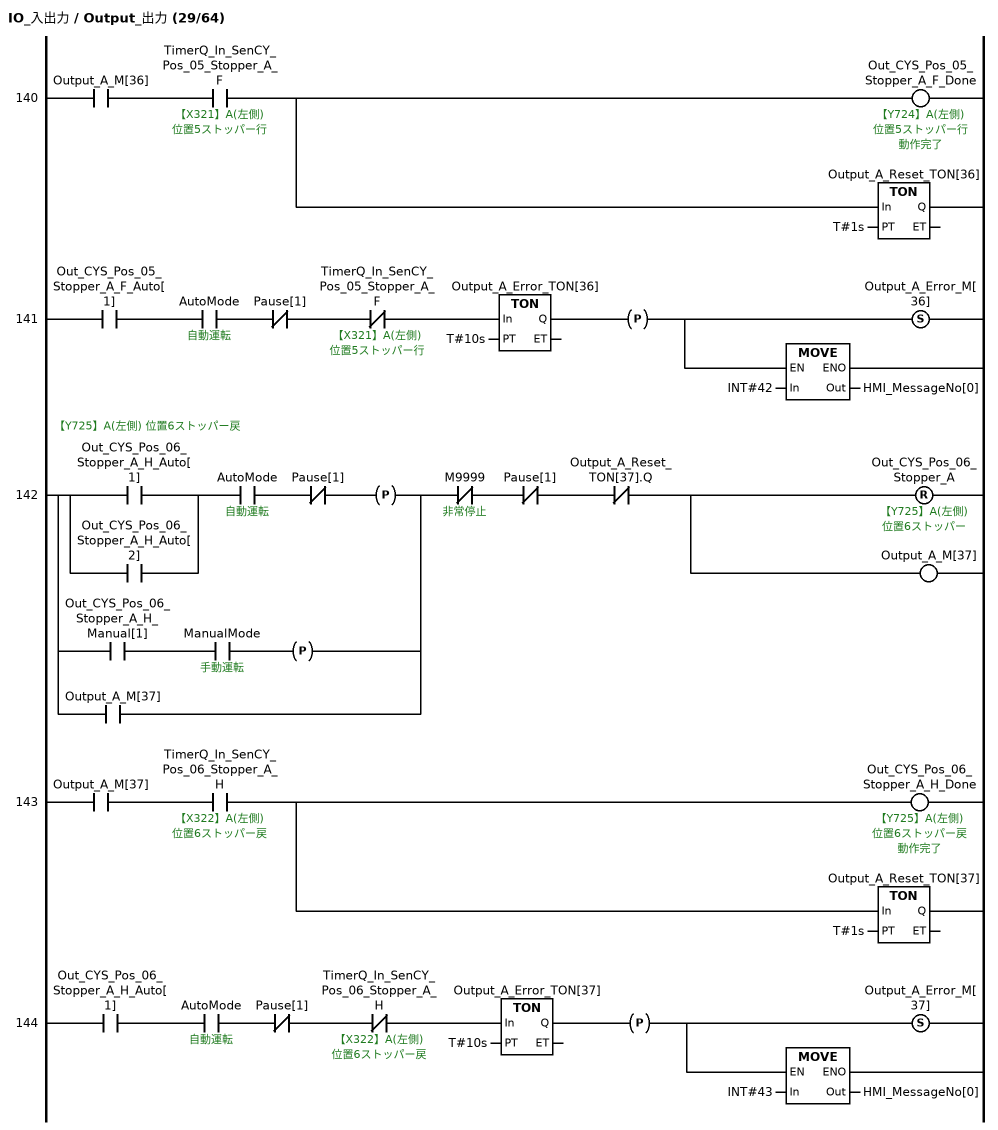
(* [picture p141: IO_入出力 / Output_出力, rungs 140-144] *)
(* Rung 140 *)
_p196 := Output_A_M[36] AND TimerQ_In_SenCY_Pos_05_Stopper_A_F;
Out_CYS_Pos_05_Stopper_A_F_Done := _p196;
Output_A_Reset_TON[36](In := _p196, PT := T#1s);
(* Rung 141 *)
Output_A_Error_TON[36](In := Out_CYS_Pos_05_Stopper_A_F_Auto[1] AND AutoMode AND NOT Pause[1] AND NOT TimerQ_In_SenCY_Pos_05_Stopper_A_F, PT := T#10s);
_e197(CLK := Output_A_Error_TON[36].Q);
IF _e197.Q THEN
    Output_A_Error_M[36] := TRUE;
    HMI_MessageNo[0] := INT#42;
END_IF;
(* Rung 142: 【Y725】A(左側) 位置6ストッパー戻 *)
_e198(CLK := (Out_CYS_Pos_06_Stopper_A_H_Auto[1] OR Out_CYS_Pos_06_Stopper_A_H_Auto[2]) AND AutoMode AND NOT Pause[1]);
_e199(CLK := Out_CYS_Pos_06_Stopper_A_H_Manual[1] AND ManualMode);
_p200 := (_e198.Q OR _e199.Q OR Output_A_M[37]) AND NOT M9999 AND NOT Pause[1] AND NOT Output_A_Reset_TON[37].Q;
IF _p200 THEN Out_CYS_Pos_06_Stopper_A := FALSE; END_IF;
Output_A_M[37] := _p200;
(* Rung 143 *)
_p201 := Output_A_M[37] AND TimerQ_In_SenCY_Pos_06_Stopper_A_H;
Out_CYS_Pos_06_Stopper_A_H_Done := _p201;
Output_A_Reset_TON[37](In := _p201, PT := T#1s);
(* Rung 144 *)
Output_A_Error_TON[37](In := Out_CYS_Pos_06_Stopper_A_H_Auto[1] AND AutoMode AND NOT Pause[1] AND NOT TimerQ_In_SenCY_Pos_06_Stopper_A_H, PT := T#10s);
_e202(CLK := Output_A_Error_TON[37].Q);
IF _e202.Q THEN
    Output_A_Error_M[37] := TRUE;
    HMI_MessageNo[0] := INT#43;
END_IF;

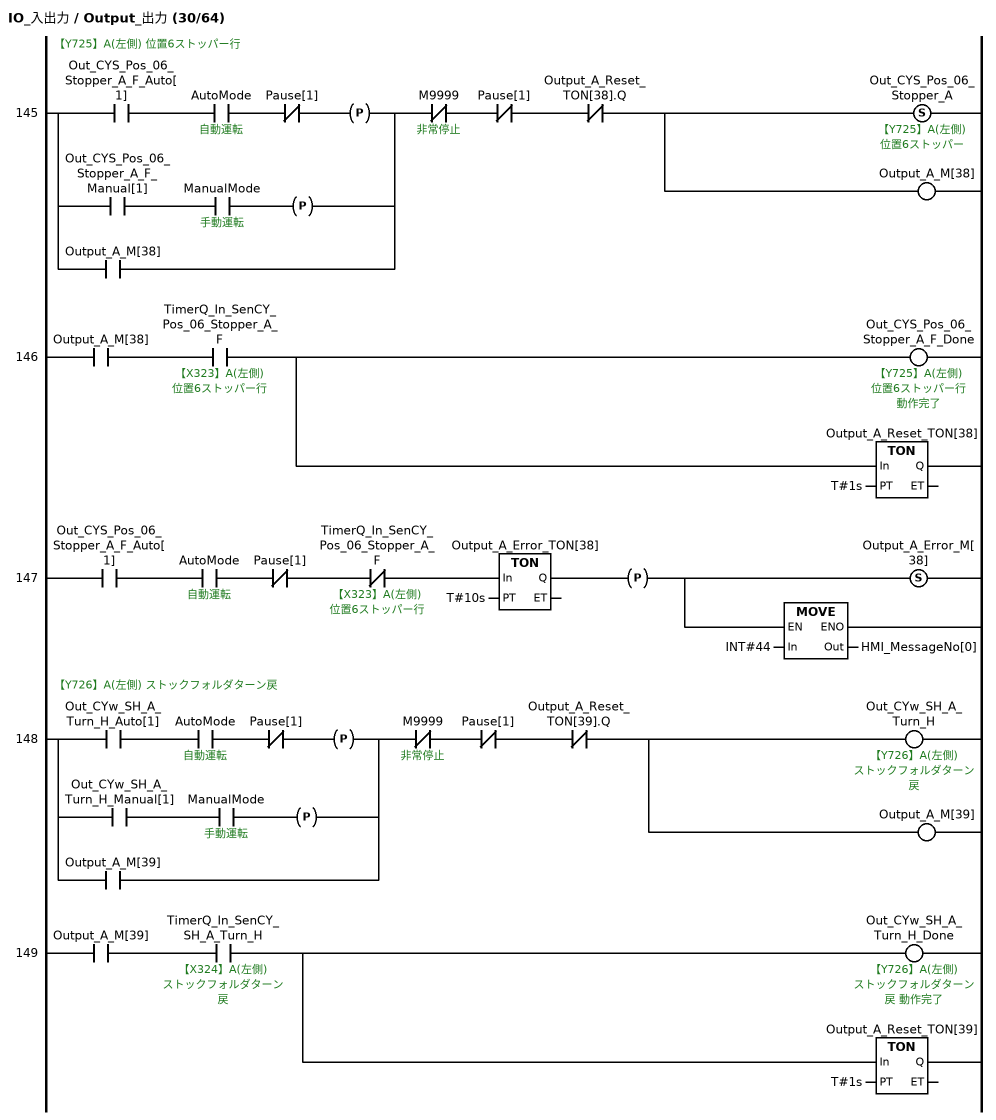
(* Rung 145: 【Y725】A(左側) 位置6ストッパー行 *)
_e203(CLK := Out_CYS_Pos_06_Stopper_A_F_Auto[1] AND AutoMode AND NOT Pause[1]);
_e204(CLK := Out_CYS_Pos_06_Stopper_A_F_Manual[1] AND ManualMode);
_p205 := (_e203.Q OR _e204.Q OR Output_A_M[38]) AND NOT M9999 AND NOT Pause[1] AND NOT Output_A_Reset_TON[38].Q;
IF _p205 THEN Out_CYS_Pos_06_Stopper_A := TRUE; END_IF;
Output_A_M[38] := _p205;
(* Rung 146 *)
_p206 := Output_A_M[38] AND TimerQ_In_SenCY_Pos_06_Stopper_A_F;
Out_CYS_Pos_06_Stopper_A_F_Done := _p206;
Output_A_Reset_TON[38](In := _p206, PT := T#1s);
(* Rung 147 *)
Output_A_Error_TON[38](In := Out_CYS_Pos_06_Stopper_A_F_Auto[1] AND AutoMode AND NOT Pause[1] AND NOT TimerQ_In_SenCY_Pos_06_Stopper_A_F, PT := T#10s);
_e207(CLK := Output_A_Error_TON[38].Q);
IF _e207.Q THEN
    Output_A_Error_M[38] := TRUE;
    HMI_MessageNo[0] := INT#44;
END_IF;
(* Rung 148: 【Y726】A(左側) ストックフォルダターン戻 *)
_e208(CLK := Out_CYw_SH_A_Turn_H_Auto[1] AND AutoMode AND NOT Pause[1]);
_e209(CLK := Out_CYw_SH_A_Turn_H_Manual[1] AND ManualMode);
_p210 := (_e208.Q OR _e209.Q OR Output_A_M[39]) AND NOT M9999 AND NOT Pause[1] AND NOT Output_A_Reset_TON[39].Q;
Out_CYw_SH_A_Turn_H := _p210;
Output_A_M[39] := _p210;
(* Rung 149 *)
Out_CYw_SH_A_Turn_H_Done := Output_A_M[39] AND TimerQ_In_SenCY_SH_A_Turn_H;
Output_A_Reset_TON[39](In := Output_A_M[39] AND TimerQ_In_SenCY_SH_A_Turn_H, PT := T#1s);

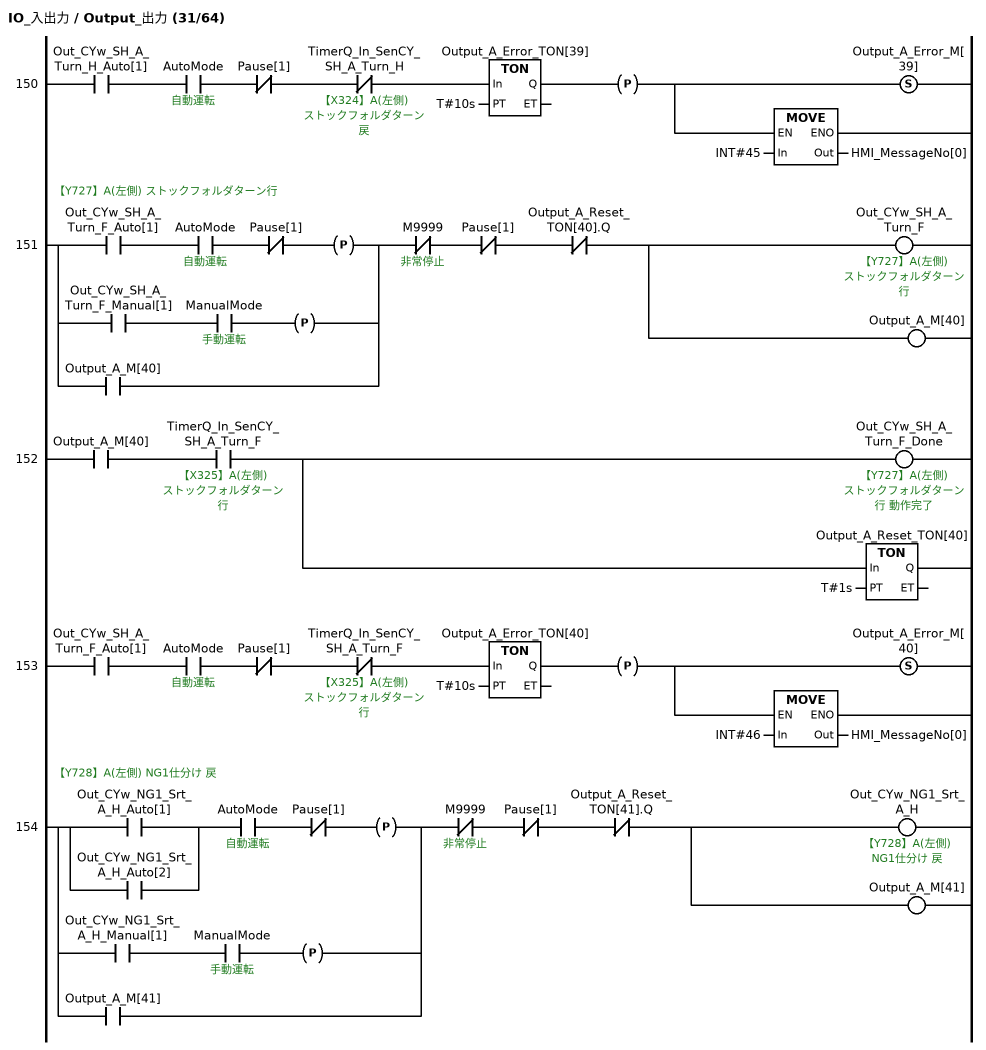
(* Rung 150 *)
Output_A_Error_TON[39](In := Out_CYw_SH_A_Turn_H_Auto[1] AND AutoMode AND NOT Pause[1] AND NOT TimerQ_In_SenCY_SH_A_Turn_H, PT := T#10s);
_e211(CLK := Output_A_Error_TON[39].Q);
IF _e211.Q THEN
    Output_A_Error_M[39] := TRUE;
    HMI_MessageNo[0] := INT#45;
END_IF;
(* Rung 151: 【Y727】A(左側) ストックフォルダターン行 *)
_e212(CLK := Out_CYw_SH_A_Turn_F_Auto[1] AND AutoMode AND NOT Pause[1]);
_e213(CLK := Out_CYw_SH_A_Turn_F_Manual[1] AND ManualMode);
_p214 := (_e212.Q OR _e213.Q OR Output_A_M[40]) AND NOT M9999 AND NOT Pause[1] AND NOT Output_A_Reset_TON[40].Q;
Out_CYw_SH_A_Turn_F := _p214;
Output_A_M[40] := _p214;
(* Rung 152 *)
Out_CYw_SH_A_Turn_F_Done := Output_A_M[40] AND TimerQ_In_SenCY_SH_A_Turn_F;
Output_A_Reset_TON[40](In := Output_A_M[40] AND TimerQ_In_SenCY_SH_A_Turn_F, PT := T#1s);
(* Rung 153 *)
Output_A_Error_TON[40](In := Out_CYw_SH_A_Turn_F_Auto[1] AND AutoMode AND NOT Pause[1] AND NOT TimerQ_In_SenCY_SH_A_Turn_F, PT := T#10s);
_e215(CLK := Output_A_Error_TON[40].Q);
IF _e215.Q THEN
    Output_A_Error_M[40] := TRUE;
    HMI_MessageNo[0] := INT#46;
END_IF;
(* Rung 154: 【Y728】A(左側) NG1仕分け 戻 *)
_e216(CLK := (Out_CYw_NG1_Srt_A_H_Auto[1] OR Out_CYw_NG1_Srt_A_H_Auto[2]) AND AutoMode AND NOT Pause[1]);
_e217(CLK := Out_CYw_NG1_Srt_A_H_Manual[1] AND ManualMode);
_p218 := (_e216.Q OR _e217.Q OR Output_A_M[41]) AND NOT M9999 AND NOT Pause[1] AND NOT Output_A_Reset_TON[41].Q;
Out_CYw_NG1_Srt_A_H := _p218;
Output_A_M[41] := _p218;

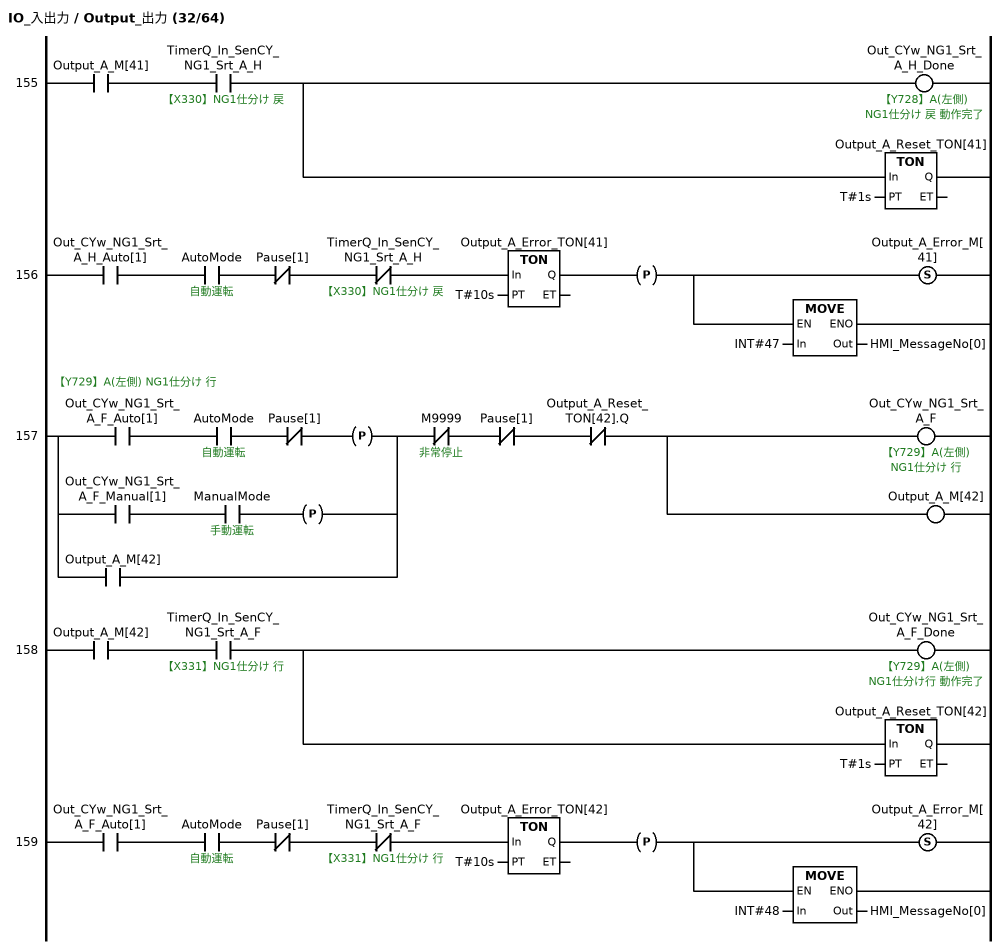
(* Rung 155 *)
Out_CYw_NG1_Srt_A_H_Done := Output_A_M[41] AND TimerQ_In_SenCY_NG1_Srt_A_H;
Output_A_Reset_TON[41](In := Output_A_M[41] AND TimerQ_In_SenCY_NG1_Srt_A_H, PT := T#1s);
(* Rung 156 *)
Output_A_Error_TON[41](In := Out_CYw_NG1_Srt_A_H_Auto[1] AND AutoMode AND NOT Pause[1] AND NOT TimerQ_In_SenCY_NG1_Srt_A_H, PT := T#10s);
_e219(CLK := Output_A_Error_TON[41].Q);
IF _e219.Q THEN
    Output_A_Error_M[41] := TRUE;
    HMI_MessageNo[0] := INT#47;
END_IF;
(* Rung 157: 【Y729】A(左側) NG1仕分け 行 *)
_e220(CLK := Out_CYw_NG1_Srt_A_F_Auto[1] AND AutoMode AND NOT Pause[1]);
_e221(CLK := Out_CYw_NG1_Srt_A_F_Manual[1] AND ManualMode);
_p222 := (_e220.Q OR _e221.Q OR Output_A_M[42]) AND NOT M9999 AND NOT Pause[1] AND NOT Output_A_Reset_TON[42].Q;
Out_CYw_NG1_Srt_A_F := _p222;
Output_A_M[42] := _p222;
(* Rung 158 *)
Out_CYw_NG1_Srt_A_F_Done := Output_A_M[42] AND TimerQ_In_SenCY_NG1_Srt_A_F;
Output_A_Reset_TON[42](In := Output_A_M[42] AND TimerQ_In_SenCY_NG1_Srt_A_F, PT := T#1s);
(* Rung 159 *)
Output_A_Error_TON[42](In := Out_CYw_NG1_Srt_A_F_Auto[1] AND AutoMode AND NOT Pause[1] AND NOT TimerQ_In_SenCY_NG1_Srt_A_F, PT := T#10s);
_e223(CLK := Output_A_Error_TON[42].Q);
IF _e223.Q THEN
    Output_A_Error_M[42] := TRUE;
    HMI_MessageNo[0] := INT#48;
END_IF;

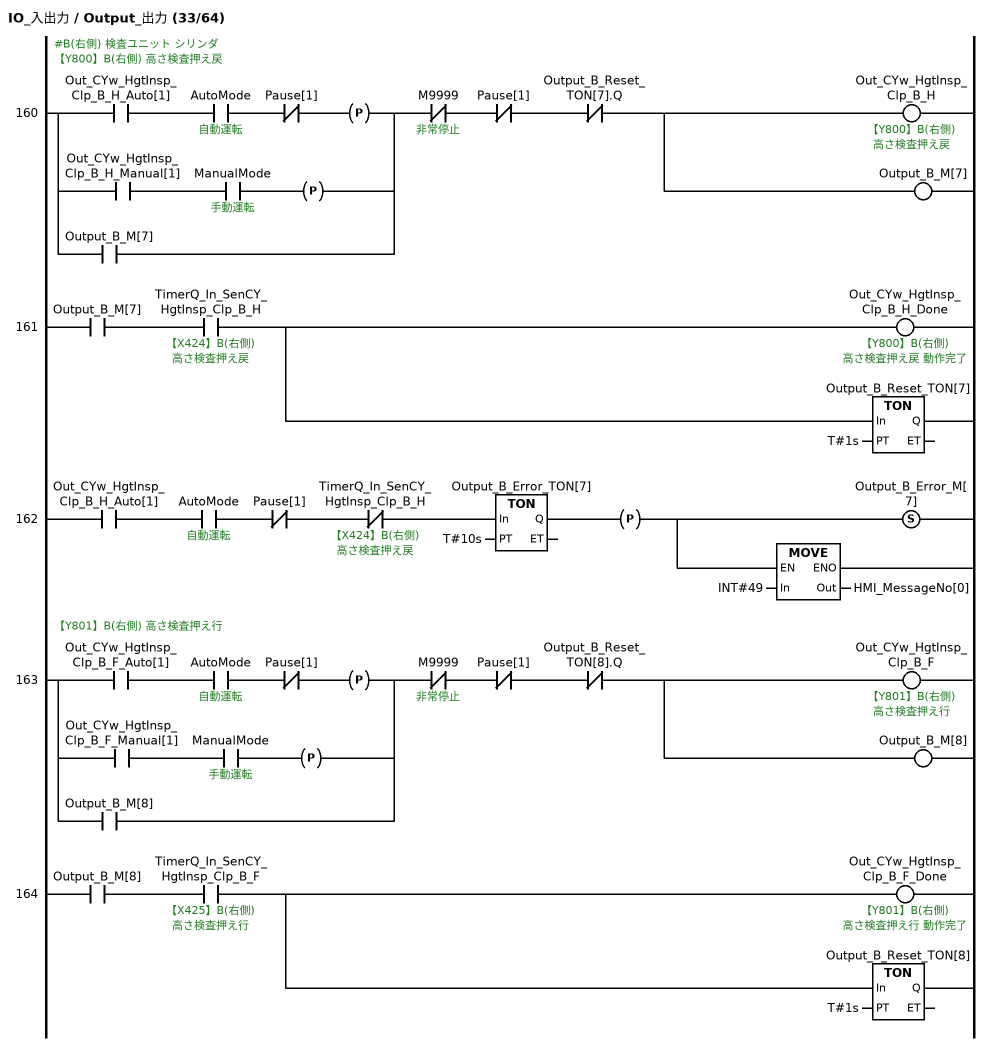
(* Rung 160: #B(右側) 検査ユニット シリンダ / 【Y800】B(右側) 高さ検査押え戻 *)
_e224(CLK := Out_CYw_HgtInsp_Clp_B_H_Auto[1] AND AutoMode AND NOT Pause[1]);
_e225(CLK := Out_CYw_HgtInsp_Clp_B_H_Manual[1] AND ManualMode);
_p226 := (_e224.Q OR _e225.Q OR Output_B_M[7]) AND NOT M9999 AND NOT Pause[1] AND NOT Output_B_Reset_TON[7].Q;
Out_CYw_HgtInsp_Clp_B_H := _p226;
Output_B_M[7] := _p226;
(* Rung 161 *)
_p227 := Output_B_M[7] AND TimerQ_In_SenCY_HgtInsp_Clp_B_H;
Out_CYw_HgtInsp_Clp_B_H_Done := _p227;
Output_B_Reset_TON[7](In := _p227, PT := T#1s);
(* Rung 162 *)
Output_B_Error_TON[7](In := Out_CYw_HgtInsp_Clp_B_H_Auto[1] AND AutoMode AND NOT Pause[1] AND NOT TimerQ_In_SenCY_HgtInsp_Clp_B_H, PT := T#10s);
_e228(CLK := Output_B_Error_TON[7].Q);
IF _e228.Q THEN
    Output_B_Error_M[7] := TRUE;
    HMI_MessageNo[0] := INT#49;
END_IF;
(* Rung 163: 【Y801】B(右側) 高さ検査押え行 *)
_e229(CLK := Out_CYw_HgtInsp_Clp_B_F_Auto[1] AND AutoMode AND NOT Pause[1]);
_e230(CLK := Out_CYw_HgtInsp_Clp_B_F_Manual[1] AND ManualMode);
_p231 := (_e229.Q OR _e230.Q OR Output_B_M[8]) AND NOT M9999 AND NOT Pause[1] AND NOT Output_B_Reset_TON[8].Q;
Out_CYw_HgtInsp_Clp_B_F := _p231;
Output_B_M[8] := _p231;
(* Rung 164 *)
_p232 := Output_B_M[8] AND TimerQ_In_SenCY_HgtInsp_Clp_B_F;
Out_CYw_HgtInsp_Clp_B_F_Done := _p232;
Output_B_Reset_TON[8](In := _p232, PT := T#1s);

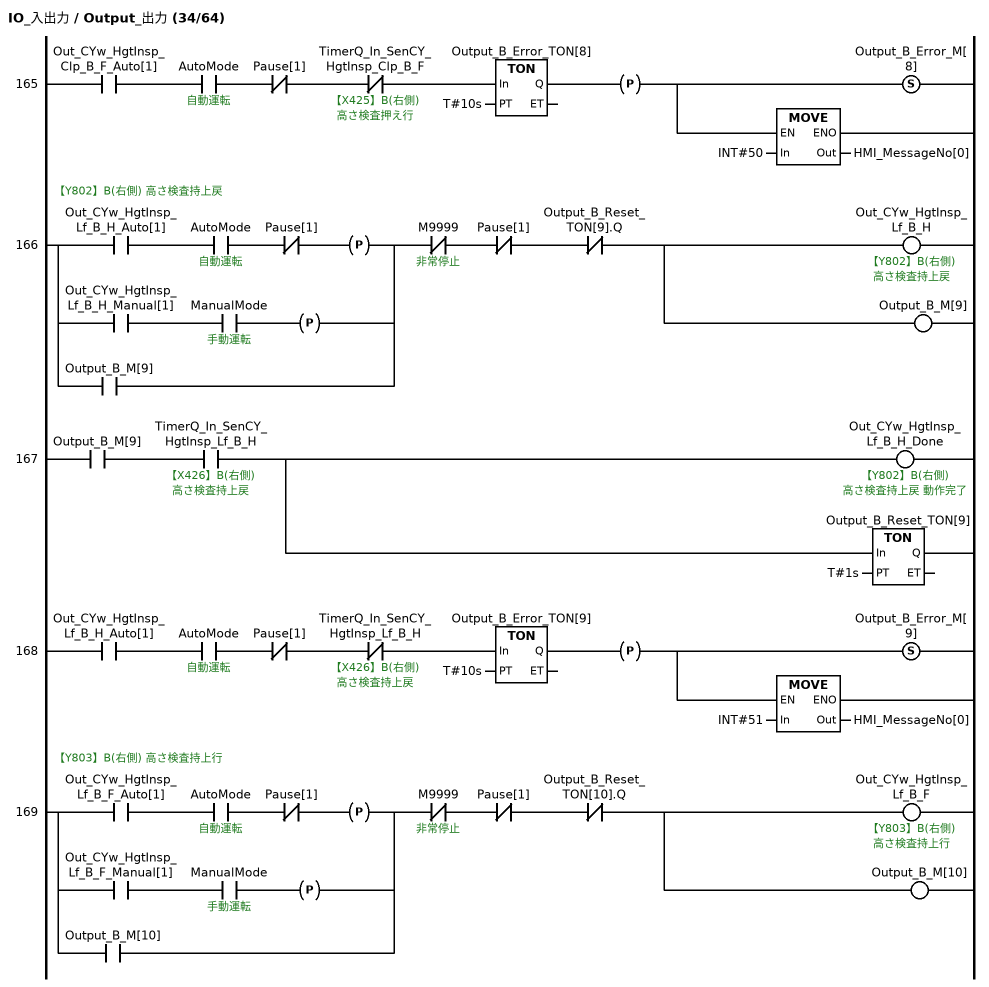
(* Rung 165 *)
Output_B_Error_TON[8](In := Out_CYw_HgtInsp_Clp_B_F_Auto[1] AND AutoMode AND NOT Pause[1] AND NOT TimerQ_In_SenCY_HgtInsp_Clp_B_F, PT := T#10s);
_e233(CLK := Output_B_Error_TON[8].Q);
IF _e233.Q THEN
    Output_B_Error_M[8] := TRUE;
    HMI_MessageNo[0] := INT#50;
END_IF;
(* Rung 166: 【Y802】B(右側) 高さ検査持上戻 *)
_e234(CLK := Out_CYw_HgtInsp_Lf_B_H_Auto[1] AND AutoMode AND NOT Pause[1]);
_e235(CLK := Out_CYw_HgtInsp_Lf_B_H_Manual[1] AND ManualMode);
_p236 := (_e234.Q OR _e235.Q OR Output_B_M[9]) AND NOT M9999 AND NOT Pause[1] AND NOT Output_B_Reset_TON[9].Q;
Out_CYw_HgtInsp_Lf_B_H := _p236;
Output_B_M[9] := _p236;
(* Rung 167 *)
Out_CYw_HgtInsp_Lf_B_H_Done := Output_B_M[9] AND TimerQ_In_SenCY_HgtInsp_Lf_B_H;
Output_B_Reset_TON[9](In := Output_B_M[9] AND TimerQ_In_SenCY_HgtInsp_Lf_B_H, PT := T#1s);
(* Rung 168 *)
Output_B_Error_TON[9](In := Out_CYw_HgtInsp_Lf_B_H_Auto[1] AND AutoMode AND NOT Pause[1] AND NOT TimerQ_In_SenCY_HgtInsp_Lf_B_H, PT := T#10s);
_e237(CLK := Output_B_Error_TON[9].Q);
IF _e237.Q THEN
    Output_B_Error_M[9] := TRUE;
    HMI_MessageNo[0] := INT#51;
END_IF;
(* Rung 169: 【Y803】B(右側) 高さ検査持上行 *)
_e238(CLK := Out_CYw_HgtInsp_Lf_B_F_Auto[1] AND AutoMode AND NOT Pause[1]);
_e239(CLK := Out_CYw_HgtInsp_Lf_B_F_Manual[1] AND ManualMode);
_p240 := (_e238.Q OR _e239.Q OR Output_B_M[10]) AND NOT M9999 AND NOT Pause[1] AND NOT Output_B_Reset_TON[10].Q;
Out_CYw_HgtInsp_Lf_B_F := _p240;
Output_B_M[10] := _p240;

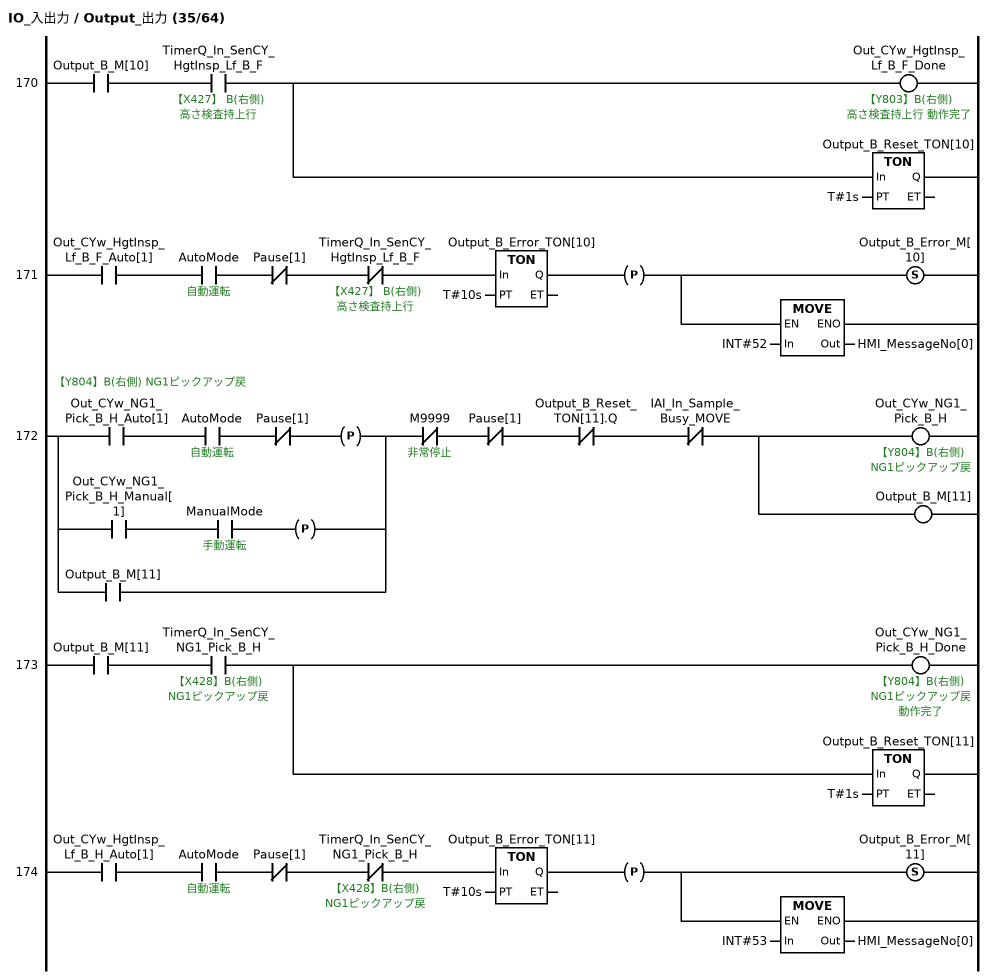
(* Rung 170 *)
_p241 := Output_B_M[10] AND TimerQ_In_SenCY_HgtInsp_Lf_B_F;
Out_CYw_HgtInsp_Lf_B_F_Done := _p241;
Output_B_Reset_TON[10](In := _p241, PT := T#1s);
(* Rung 171 *)
Output_B_Error_TON[10](In := Out_CYw_HgtInsp_Lf_B_F_Auto[1] AND AutoMode AND NOT Pause[1] AND NOT TimerQ_In_SenCY_HgtInsp_Lf_B_F, PT := T#10s);
_e242(CLK := Output_B_Error_TON[10].Q);
IF _e242.Q THEN
    Output_B_Error_M[10] := TRUE;
    HMI_MessageNo[0] := INT#52;
END_IF;
(* Rung 172: 【Y804】B(右側) NG1ピックアップ戻 *)
_e243(CLK := Out_CYw_NG1_Pick_B_H_Auto[1] AND AutoMode AND NOT Pause[1]);
_e244(CLK := Out_CYw_NG1_Pick_B_H_Manual[1] AND ManualMode);
_p245 := (_e243.Q OR _e244.Q OR Output_B_M[11]) AND NOT M9999 AND NOT Pause[1] AND NOT Output_B_Reset_TON[11].Q AND NOT IAI_In_Sample_Busy_MOVE;
Out_CYw_NG1_Pick_B_H := _p245;
Output_B_M[11] := _p245;
(* Rung 173 *)
Out_CYw_NG1_Pick_B_H_Done := Output_B_M[11] AND TimerQ_In_SenCY_NG1_Pick_B_H;
Output_B_Reset_TON[11](In := Output_B_M[11] AND TimerQ_In_SenCY_NG1_Pick_B_H, PT := T#1s);
(* Rung 174 *)
Output_B_Error_TON[11](In := Out_CYw_HgtInsp_Lf_B_H_Auto[1] AND AutoMode AND NOT Pause[1] AND NOT TimerQ_In_SenCY_NG1_Pick_B_H, PT := T#10s);
_e246(CLK := Output_B_Error_TON[11].Q);
IF _e246.Q THEN
    Output_B_Error_M[11] := TRUE;
    HMI_MessageNo[0] := INT#53;
END_IF;

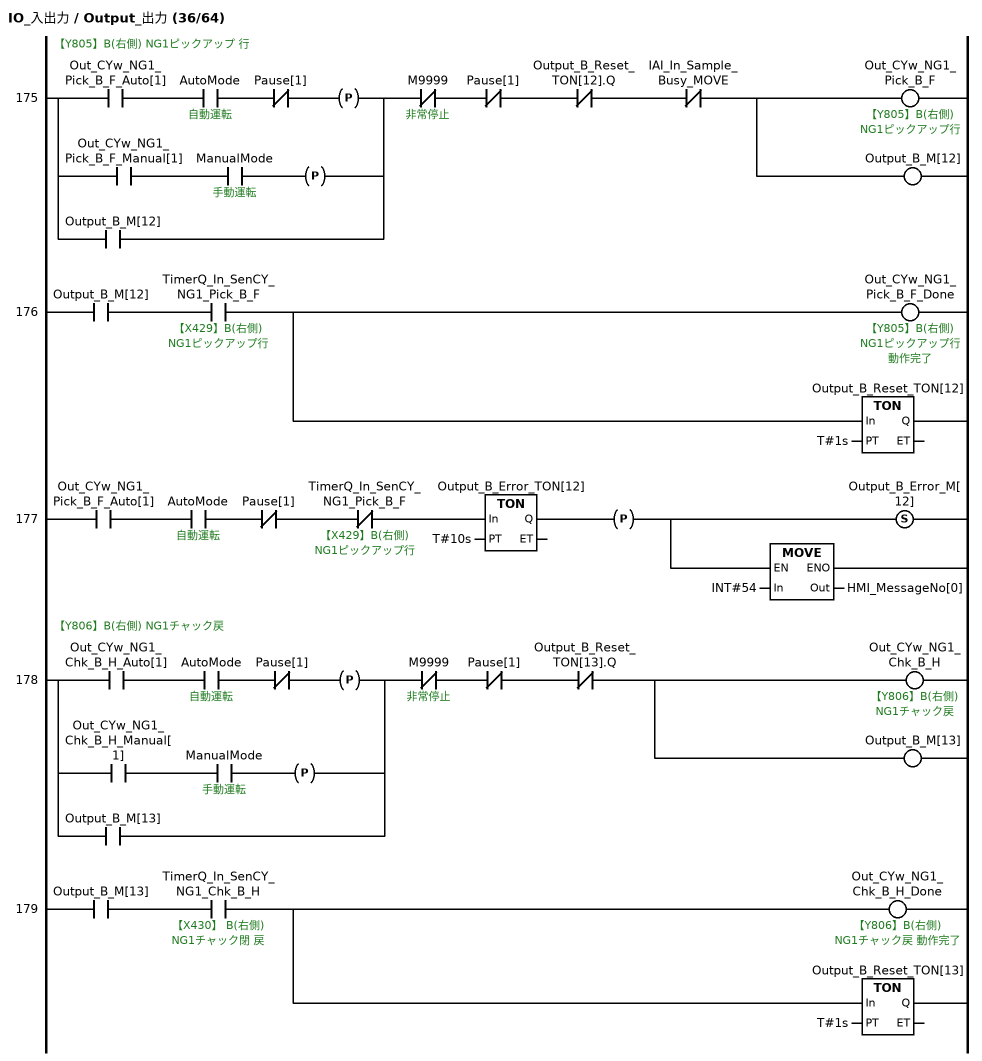
(* Rung 175: 【Y805】B(右側) NG1ピックアップ 行 *)
_e247(CLK := Out_CYw_NG1_Pick_B_F_Auto[1] AND AutoMode AND NOT Pause[1]);
_e248(CLK := Out_CYw_NG1_Pick_B_F_Manual[1] AND ManualMode);
_p249 := (_e247.Q OR _e248.Q OR Output_B_M[12]) AND NOT M9999 AND NOT Pause[1] AND NOT Output_B_Reset_TON[12].Q AND NOT IAI_In_Sample_Busy_MOVE;
Out_CYw_NG1_Pick_B_F := _p249;
Output_B_M[12] := _p249;
(* Rung 176 *)
Out_CYw_NG1_Pick_B_F_Done := Output_B_M[12] AND TimerQ_In_SenCY_NG1_Pick_B_F;
Output_B_Reset_TON[12](In := Output_B_M[12] AND TimerQ_In_SenCY_NG1_Pick_B_F, PT := T#1s);
(* Rung 177 *)
Output_B_Error_TON[12](In := Out_CYw_NG1_Pick_B_F_Auto[1] AND AutoMode AND NOT Pause[1] AND NOT TimerQ_In_SenCY_NG1_Pick_B_F, PT := T#10s);
_e250(CLK := Output_B_Error_TON[12].Q);
IF _e250.Q THEN
    Output_B_Error_M[12] := TRUE;
    HMI_MessageNo[0] := INT#54;
END_IF;
(* Rung 178: 【Y806】B(右側) NG1チャック戻 *)
_e251(CLK := Out_CYw_NG1_Chk_B_H_Auto[1] AND AutoMode AND NOT Pause[1]);
_e252(CLK := Out_CYw_NG1_Chk_B_H_Manual[1] AND ManualMode);
_p253 := (_e251.Q OR _e252.Q OR Output_B_M[13]) AND NOT M9999 AND NOT Pause[1] AND NOT Output_B_Reset_TON[13].Q;
Out_CYw_NG1_Chk_B_H := _p253;
Output_B_M[13] := _p253;
(* Rung 179 *)
Out_CYw_NG1_Chk_B_H_Done := Output_B_M[13] AND TimerQ_In_SenCY_NG1_Chk_B_H;
Output_B_Reset_TON[13](In := Output_B_M[13] AND TimerQ_In_SenCY_NG1_Chk_B_H, PT := T#1s);

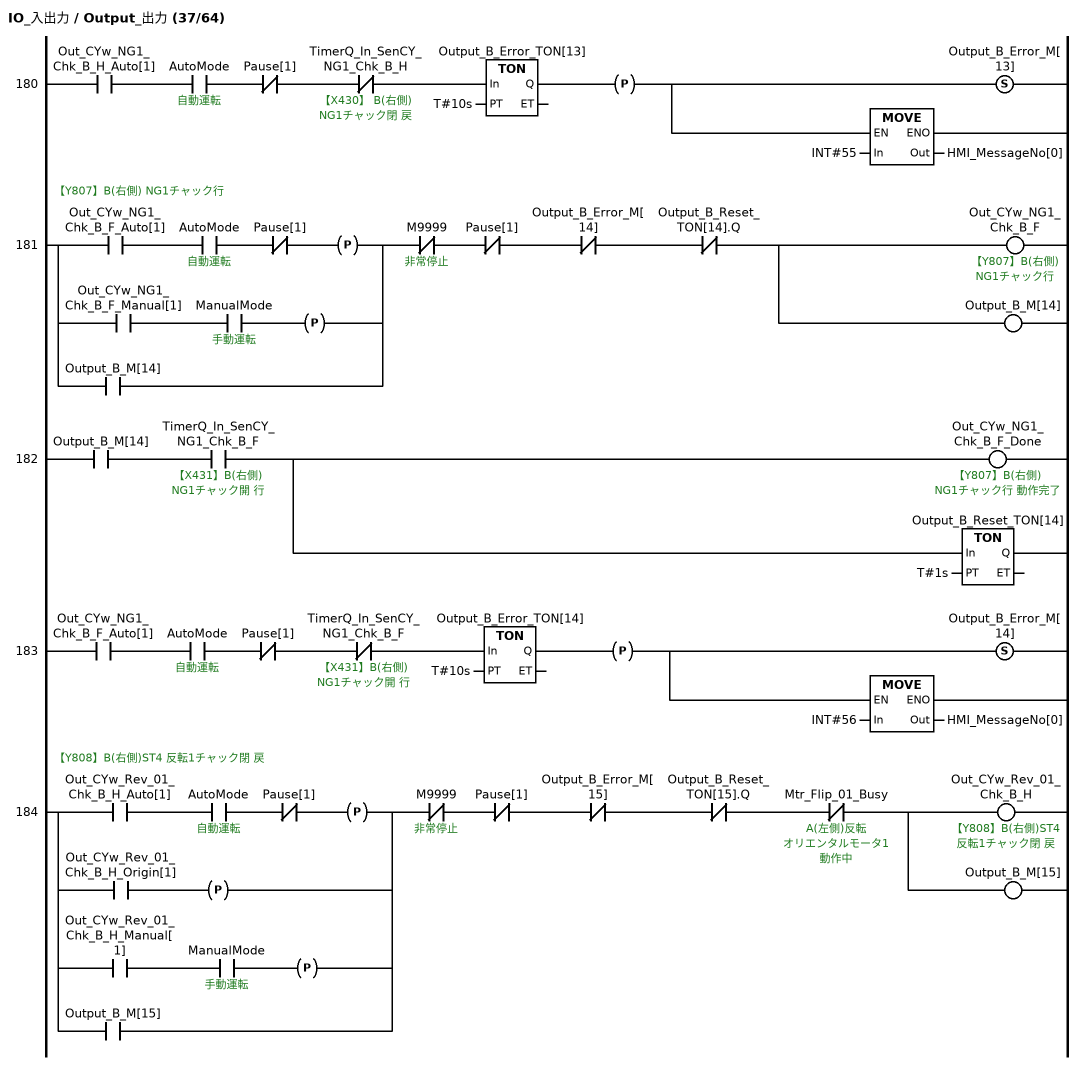
(* Rung 180 *)
Output_B_Error_TON[13](In := Out_CYw_NG1_Chk_B_H_Auto[1] AND AutoMode AND NOT Pause[1] AND NOT TimerQ_In_SenCY_NG1_Chk_B_H, PT := T#10s);
_e254(CLK := Output_B_Error_TON[13].Q);
IF _e254.Q THEN
    Output_B_Error_M[13] := TRUE;
    HMI_MessageNo[0] := INT#55;
END_IF;
(* Rung 181: 【Y807】B(右側) NG1チャック行 *)
_e255(CLK := Out_CYw_NG1_Chk_B_F_Auto[1] AND AutoMode AND NOT Pause[1]);
_e256(CLK := Out_CYw_NG1_Chk_B_F_Manual[1] AND ManualMode);
_p257 := (_e255.Q OR _e256.Q OR Output_B_M[14]) AND NOT M9999 AND NOT Pause[1] AND NOT Output_B_Error_M[14] AND NOT Output_B_Reset_TON[14].Q;
Out_CYw_NG1_Chk_B_F := _p257;
Output_B_M[14] := _p257;
(* Rung 182 *)
Out_CYw_NG1_Chk_B_F_Done := Output_B_M[14] AND TimerQ_In_SenCY_NG1_Chk_B_F;
Output_B_Reset_TON[14](In := Output_B_M[14] AND TimerQ_In_SenCY_NG1_Chk_B_F, PT := T#1s);
(* Rung 183 *)
Output_B_Error_TON[14](In := Out_CYw_NG1_Chk_B_F_Auto[1] AND AutoMode AND NOT Pause[1] AND NOT TimerQ_In_SenCY_NG1_Chk_B_F, PT := T#10s);
_e258(CLK := Output_B_Error_TON[14].Q);
IF _e258.Q THEN
    Output_B_Error_M[14] := TRUE;
    HMI_MessageNo[0] := INT#56;
END_IF;
(* Rung 184: 【Y808】B(右側)ST4 反転1チャック閉 戻 *)
_e259(CLK := Out_CYw_Rev_01_Chk_B_H_Auto[1] AND AutoMode AND NOT Pause[1]);
_e260(CLK := Out_CYw_Rev_01_Chk_B_H_Origin[1]);
_e261(CLK := Out_CYw_Rev_01_Chk_B_H_Manual[1] AND ManualMode);
_p262 := (_e259.Q OR _e260.Q OR _e261.Q OR Output_B_M[15]) AND NOT M9999 AND NOT Pause[1] AND NOT Output_B_Error_M[15] AND NOT Output_B_Reset_TON[15].Q AND NOT Mtr_Flip_01_Busy;
Out_CYw_Rev_01_Chk_B_H := _p262;
Output_B_M[15] := _p262;

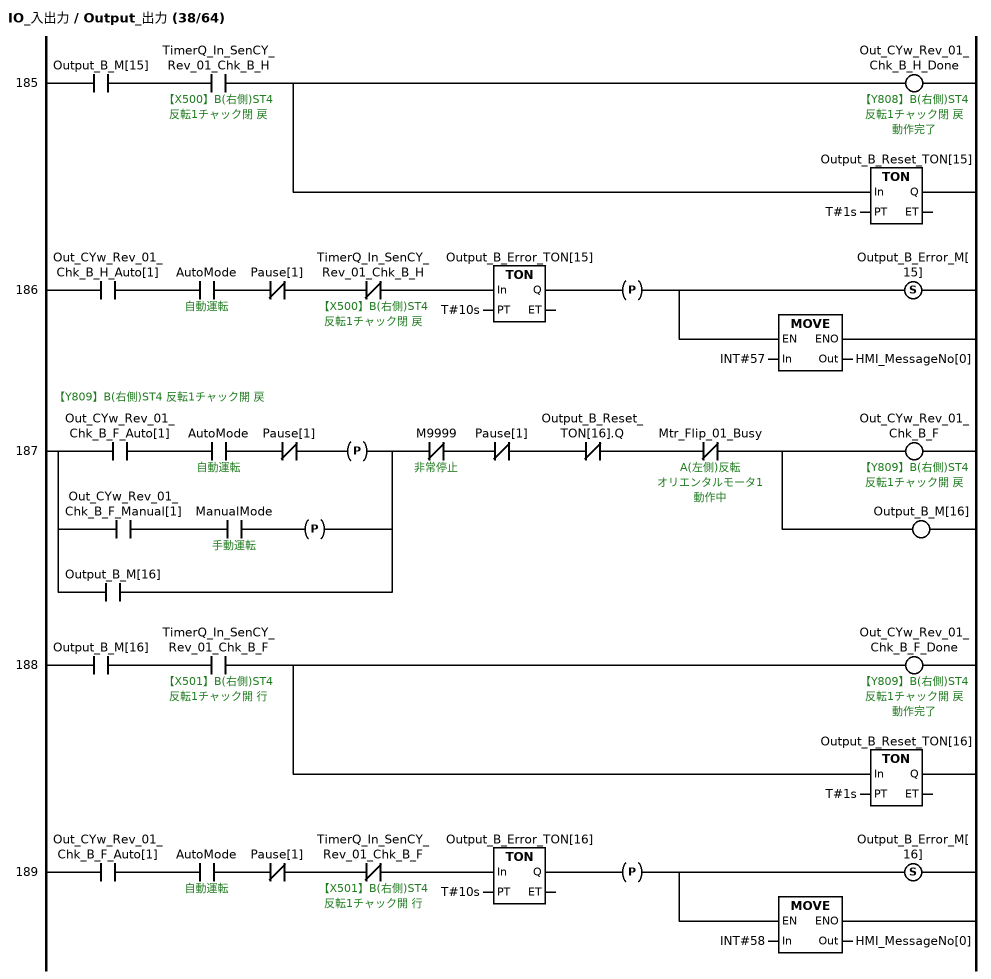
(* Rung 185 *)
_p263 := Output_B_M[15] AND TimerQ_In_SenCY_Rev_01_Chk_B_H;
Out_CYw_Rev_01_Chk_B_H_Done := _p263;
Output_B_Reset_TON[15](In := _p263, PT := T#1s);
(* Rung 186 *)
Output_B_Error_TON[15](In := Out_CYw_Rev_01_Chk_B_H_Auto[1] AND AutoMode AND NOT Pause[1] AND NOT TimerQ_In_SenCY_Rev_01_Chk_B_H, PT := T#10s);
_e264(CLK := Output_B_Error_TON[15].Q);
IF _e264.Q THEN
    Output_B_Error_M[15] := TRUE;
    HMI_MessageNo[0] := INT#57;
END_IF;
(* Rung 187: 【Y809】B(右側)ST4 反転1チャック開 戻 *)
_e265(CLK := Out_CYw_Rev_01_Chk_B_F_Auto[1] AND AutoMode AND NOT Pause[1]);
_e266(CLK := Out_CYw_Rev_01_Chk_B_F_Manual[1] AND ManualMode);
_p267 := (_e265.Q OR _e266.Q OR Output_B_M[16]) AND NOT M9999 AND NOT Pause[1] AND NOT Output_B_Reset_TON[16].Q AND NOT Mtr_Flip_01_Busy;
Out_CYw_Rev_01_Chk_B_F := _p267;
Output_B_M[16] := _p267;
(* Rung 188 *)
_p268 := Output_B_M[16] AND TimerQ_In_SenCY_Rev_01_Chk_B_F;
Out_CYw_Rev_01_Chk_B_F_Done := _p268;
Output_B_Reset_TON[16](In := _p268, PT := T#1s);
(* Rung 189 *)
Output_B_Error_TON[16](In := Out_CYw_Rev_01_Chk_B_F_Auto[1] AND AutoMode AND NOT Pause[1] AND NOT TimerQ_In_SenCY_Rev_01_Chk_B_F, PT := T#10s);
_e269(CLK := Output_B_Error_TON[16].Q);
IF _e269.Q THEN
    Output_B_Error_M[16] := TRUE;
    HMI_MessageNo[0] := INT#58;
END_IF;

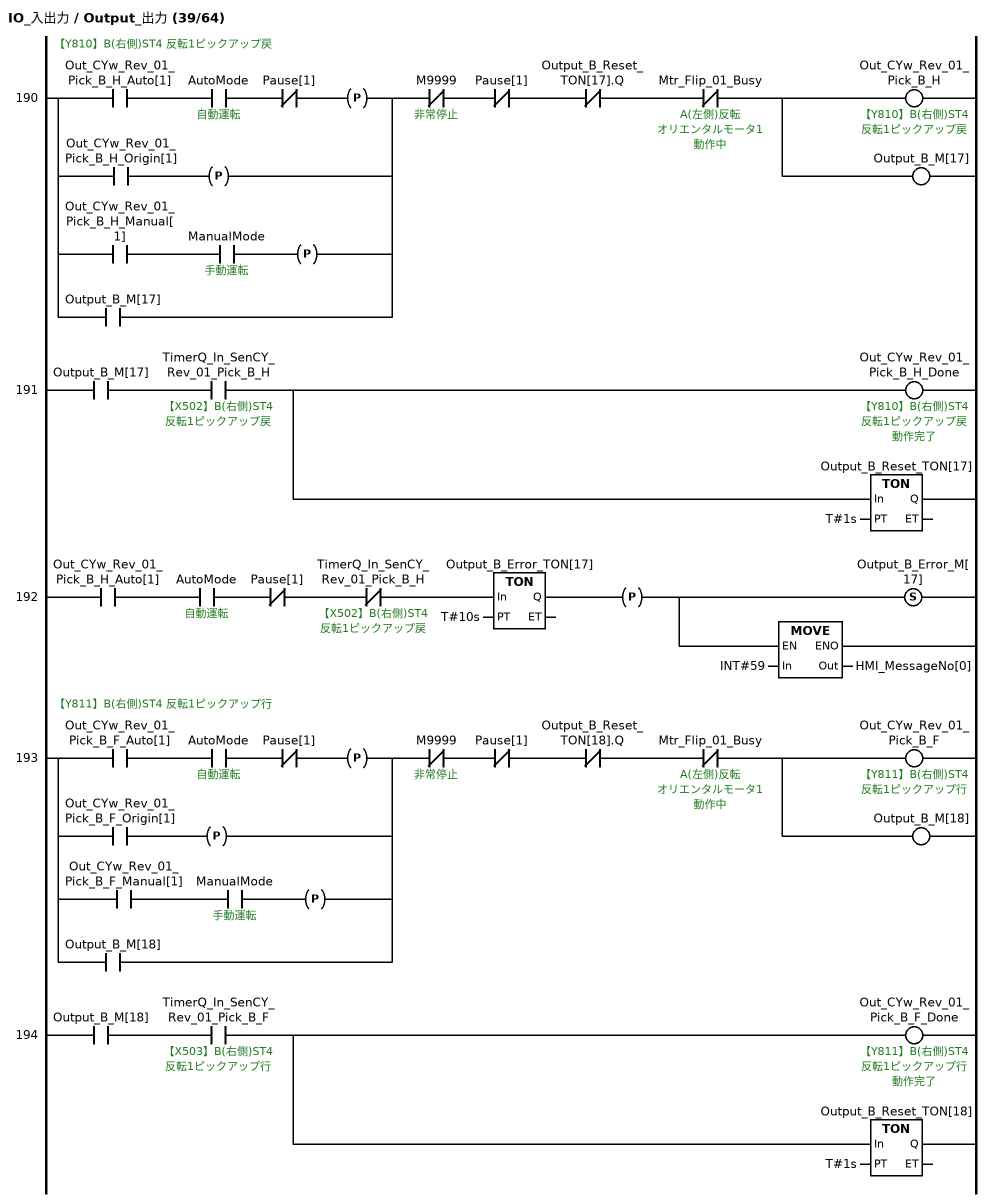
(* Rung 190: 【Y810】B(右側)ST4 反転1ピックアップ戻 *)
_e270(CLK := Out_CYw_Rev_01_Pick_B_H_Auto[1] AND AutoMode AND NOT Pause[1]);
_e271(CLK := Out_CYw_Rev_01_Pick_B_H_Origin[1]);
_e272(CLK := Out_CYw_Rev_01_Pick_B_H_Manual[1] AND ManualMode);
_p273 := (_e270.Q OR _e271.Q OR _e272.Q OR Output_B_M[17]) AND NOT M9999 AND NOT Pause[1] AND NOT Output_B_Reset_TON[17].Q AND NOT Mtr_Flip_01_Busy;
Out_CYw_Rev_01_Pick_B_H := _p273;
Output_B_M[17] := _p273;
(* Rung 191 *)
_p274 := Output_B_M[17] AND TimerQ_In_SenCY_Rev_01_Pick_B_H;
Out_CYw_Rev_01_Pick_B_H_Done := _p274;
Output_B_Reset_TON[17](In := _p274, PT := T#1s);
(* Rung 192 *)
Output_B_Error_TON[17](In := Out_CYw_Rev_01_Pick_B_H_Auto[1] AND AutoMode AND NOT Pause[1] AND NOT TimerQ_In_SenCY_Rev_01_Pick_B_H, PT := T#10s);
_e275(CLK := Output_B_Error_TON[17].Q);
IF _e275.Q THEN
    Output_B_Error_M[17] := TRUE;
    HMI_MessageNo[0] := INT#59;
END_IF;
(* Rung 193: 【Y811】B(右側)ST4 反転1ピックアップ行 *)
_e276(CLK := Out_CYw_Rev_01_Pick_B_F_Auto[1] AND AutoMode AND NOT Pause[1]);
_e277(CLK := Out_CYw_Rev_01_Pick_B_F_Origin[1]);
_e278(CLK := Out_CYw_Rev_01_Pick_B_F_Manual[1] AND ManualMode);
_p279 := (_e276.Q OR _e277.Q OR _e278.Q OR Output_B_M[18]) AND NOT M9999 AND NOT Pause[1] AND NOT Output_B_Reset_TON[18].Q AND NOT Mtr_Flip_01_Busy;
Out_CYw_Rev_01_Pick_B_F := _p279;
Output_B_M[18] := _p279;
(* Rung 194 *)
_p280 := Output_B_M[18] AND TimerQ_In_SenCY_Rev_01_Pick_B_F;
Out_CYw_Rev_01_Pick_B_F_Done := _p280;
Output_B_Reset_TON[18](In := _p280, PT := T#1s);

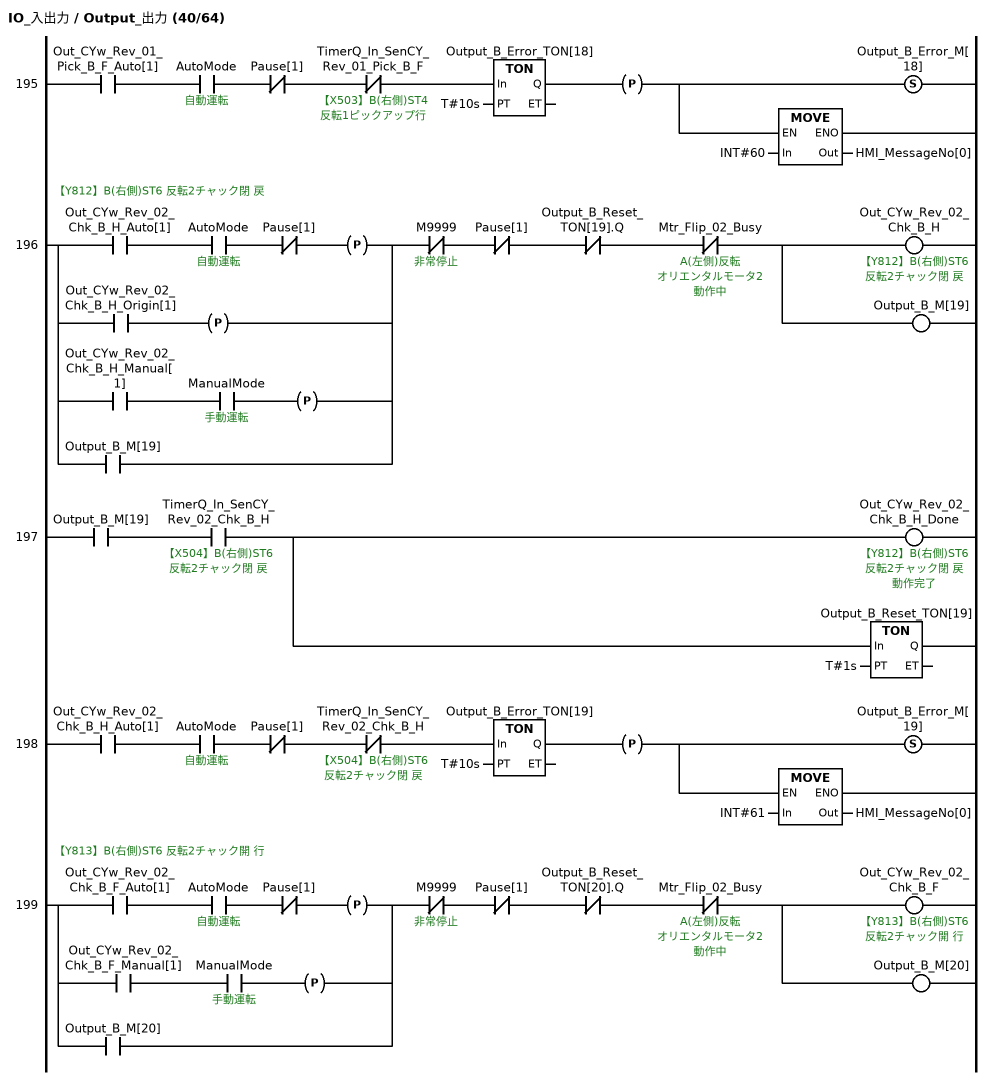
(* Rung 195 *)
Output_B_Error_TON[18](In := Out_CYw_Rev_01_Pick_B_F_Auto[1] AND AutoMode AND NOT Pause[1] AND NOT TimerQ_In_SenCY_Rev_01_Pick_B_F, PT := T#10s);
_e281(CLK := Output_B_Error_TON[18].Q);
IF _e281.Q THEN
    Output_B_Error_M[18] := TRUE;
    HMI_MessageNo[0] := INT#60;
END_IF;
(* Rung 196: 【Y812】B(右側)ST6 反転2チャック閉 戻 *)
_e282(CLK := Out_CYw_Rev_02_Chk_B_H_Auto[1] AND AutoMode AND NOT Pause[1]);
_e283(CLK := Out_CYw_Rev_02_Chk_B_H_Origin[1]);
_e284(CLK := Out_CYw_Rev_02_Chk_B_H_Manual[1] AND ManualMode);
_p285 := (_e282.Q OR _e283.Q OR _e284.Q OR Output_B_M[19]) AND NOT M9999 AND NOT Pause[1] AND NOT Output_B_Reset_TON[19].Q AND NOT Mtr_Flip_02_Busy;
Out_CYw_Rev_02_Chk_B_H := _p285;
Output_B_M[19] := _p285;
(* Rung 197 *)
_p286 := Output_B_M[19] AND TimerQ_In_SenCY_Rev_02_Chk_B_H;
Out_CYw_Rev_02_Chk_B_H_Done := _p286;
Output_B_Reset_TON[19](In := _p286, PT := T#1s);
(* Rung 198 *)
Output_B_Error_TON[19](In := Out_CYw_Rev_02_Chk_B_H_Auto[1] AND AutoMode AND NOT Pause[1] AND NOT TimerQ_In_SenCY_Rev_02_Chk_B_H, PT := T#10s);
_e287(CLK := Output_B_Error_TON[19].Q);
IF _e287.Q THEN
    Output_B_Error_M[19] := TRUE;
    HMI_MessageNo[0] := INT#61;
END_IF;
(* Rung 199: 【Y813】B(右側)ST6 反転2チャック開 行 *)
_e288(CLK := Out_CYw_Rev_02_Chk_B_F_Auto[1] AND AutoMode AND NOT Pause[1]);
_e289(CLK := Out_CYw_Rev_02_Chk_B_F_Manual[1] AND ManualMode);
_p290 := (_e288.Q OR _e289.Q OR Output_B_M[20]) AND NOT M9999 AND NOT Pause[1] AND NOT Output_B_Reset_TON[20].Q AND NOT Mtr_Flip_02_Busy;
Out_CYw_Rev_02_Chk_B_F := _p290;
Output_B_M[20] := _p290;

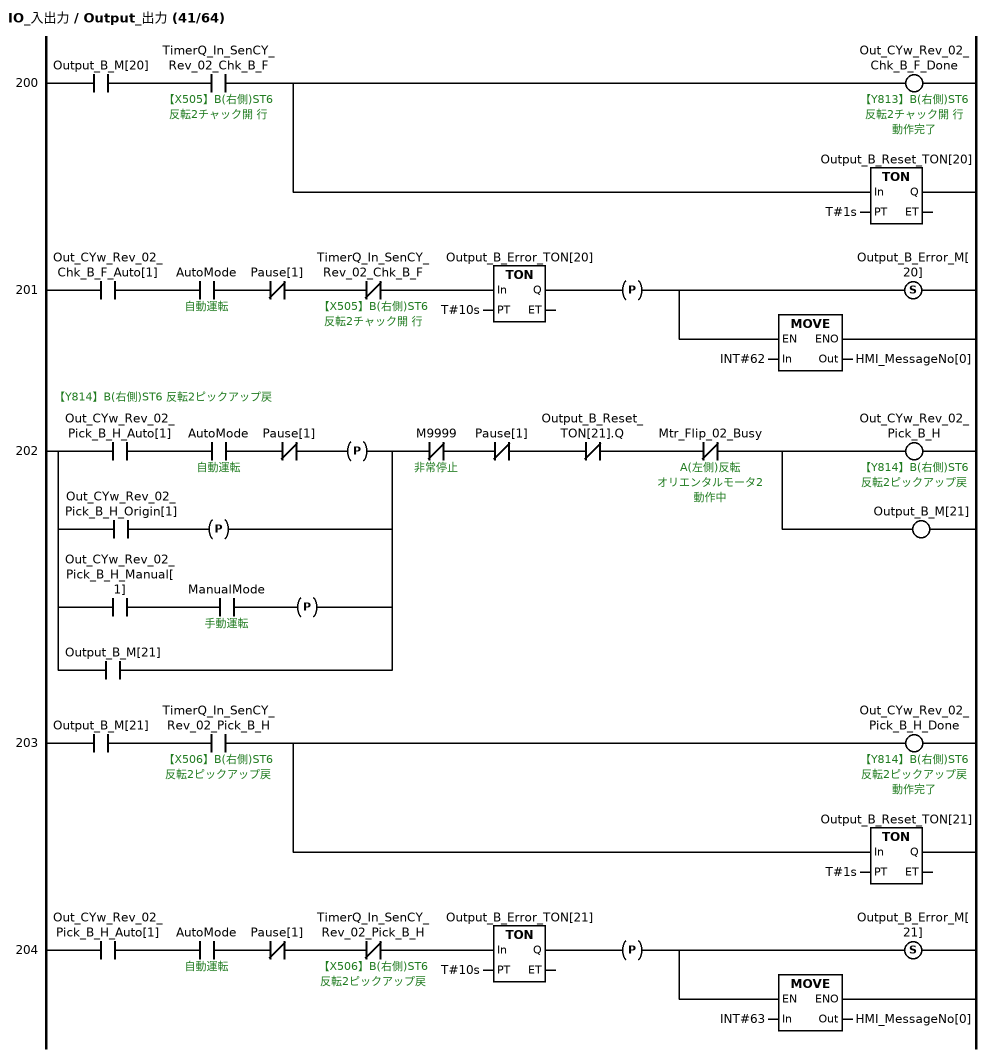
(* Rung 200 *)
_p291 := Output_B_M[20] AND TimerQ_In_SenCY_Rev_02_Chk_B_F;
Out_CYw_Rev_02_Chk_B_F_Done := _p291;
Output_B_Reset_TON[20](In := _p291, PT := T#1s);
(* Rung 201 *)
Output_B_Error_TON[20](In := Out_CYw_Rev_02_Chk_B_F_Auto[1] AND AutoMode AND NOT Pause[1] AND NOT TimerQ_In_SenCY_Rev_02_Chk_B_F, PT := T#10s);
_e292(CLK := Output_B_Error_TON[20].Q);
IF _e292.Q THEN
    Output_B_Error_M[20] := TRUE;
    HMI_MessageNo[0] := INT#62;
END_IF;
(* Rung 202: 【Y814】B(右側)ST6 反転2ピックアップ戻 *)
_e293(CLK := Out_CYw_Rev_02_Pick_B_H_Auto[1] AND AutoMode AND NOT Pause[1]);
_e294(CLK := Out_CYw_Rev_02_Pick_B_H_Origin[1]);
_e295(CLK := Out_CYw_Rev_02_Pick_B_H_Manual[1] AND ManualMode);
_p296 := (_e293.Q OR _e294.Q OR _e295.Q OR Output_B_M[21]) AND NOT M9999 AND NOT Pause[1] AND NOT Output_B_Reset_TON[21].Q AND NOT Mtr_Flip_02_Busy;
Out_CYw_Rev_02_Pick_B_H := _p296;
Output_B_M[21] := _p296;
(* Rung 203 *)
_p297 := Output_B_M[21] AND TimerQ_In_SenCY_Rev_02_Pick_B_H;
Out_CYw_Rev_02_Pick_B_H_Done := _p297;
Output_B_Reset_TON[21](In := _p297, PT := T#1s);
(* Rung 204 *)
Output_B_Error_TON[21](In := Out_CYw_Rev_02_Pick_B_H_Auto[1] AND AutoMode AND NOT Pause[1] AND NOT TimerQ_In_SenCY_Rev_02_Pick_B_H, PT := T#10s);
_e298(CLK := Output_B_Error_TON[21].Q);
IF _e298.Q THEN
    Output_B_Error_M[21] := TRUE;
    HMI_MessageNo[0] := INT#63;
END_IF;

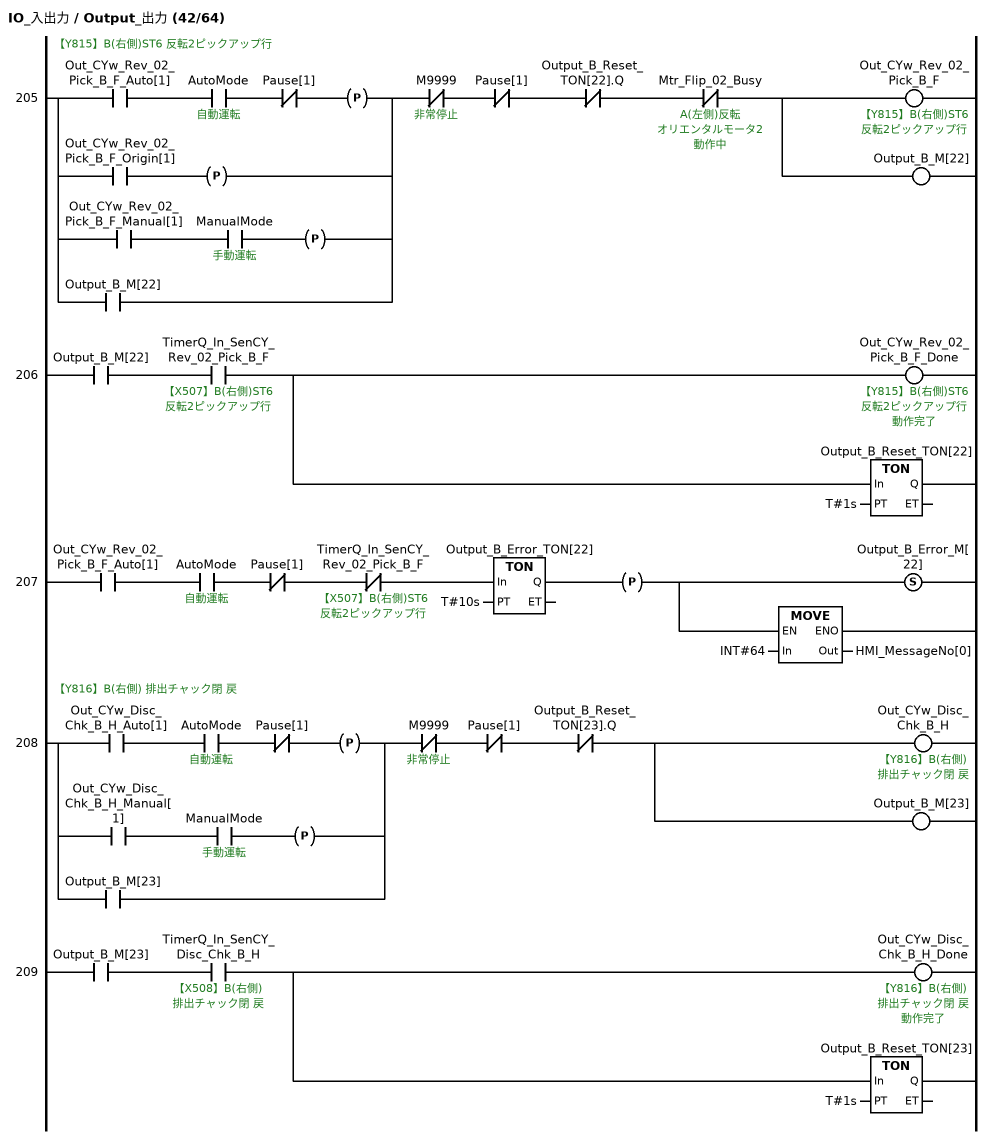
(* Rung 205: 【Y815】B(右側)ST6 反転2ピックアップ行 *)
_e299(CLK := Out_CYw_Rev_02_Pick_B_F_Auto[1] AND AutoMode AND NOT Pause[1]);
_e300(CLK := Out_CYw_Rev_02_Pick_B_F_Origin[1]);
_e301(CLK := Out_CYw_Rev_02_Pick_B_F_Manual[1] AND ManualMode);
_p302 := (_e299.Q OR _e300.Q OR _e301.Q OR Output_B_M[22]) AND NOT M9999 AND NOT Pause[1] AND NOT Output_B_Reset_TON[22].Q AND NOT Mtr_Flip_02_Busy;
Out_CYw_Rev_02_Pick_B_F := _p302;
Output_B_M[22] := _p302;
(* Rung 206 *)
_p303 := Output_B_M[22] AND TimerQ_In_SenCY_Rev_02_Pick_B_F;
Out_CYw_Rev_02_Pick_B_F_Done := _p303;
Output_B_Reset_TON[22](In := _p303, PT := T#1s);
(* Rung 207 *)
Output_B_Error_TON[22](In := Out_CYw_Rev_02_Pick_B_F_Auto[1] AND AutoMode AND NOT Pause[1] AND NOT TimerQ_In_SenCY_Rev_02_Pick_B_F, PT := T#10s);
_e304(CLK := Output_B_Error_TON[22].Q);
IF _e304.Q THEN
    Output_B_Error_M[22] := TRUE;
    HMI_MessageNo[0] := INT#64;
END_IF;
(* Rung 208: 【Y816】B(右側) 排出チャック閉 戻 *)
_e305(CLK := Out_CYw_Disc_Chk_B_H_Auto[1] AND AutoMode AND NOT Pause[1]);
_e306(CLK := Out_CYw_Disc_Chk_B_H_Manual[1] AND ManualMode);
_p307 := (_e305.Q OR _e306.Q OR Output_B_M[23]) AND NOT M9999 AND NOT Pause[1] AND NOT Output_B_Reset_TON[23].Q;
Out_CYw_Disc_Chk_B_H := _p307;
Output_B_M[23] := _p307;
(* Rung 209 *)
Out_CYw_Disc_Chk_B_H_Done := Output_B_M[23] AND TimerQ_In_SenCY_Disc_Chk_B_H;
Output_B_Reset_TON[23](In := Output_B_M[23] AND TimerQ_In_SenCY_Disc_Chk_B_H, PT := T#1s);

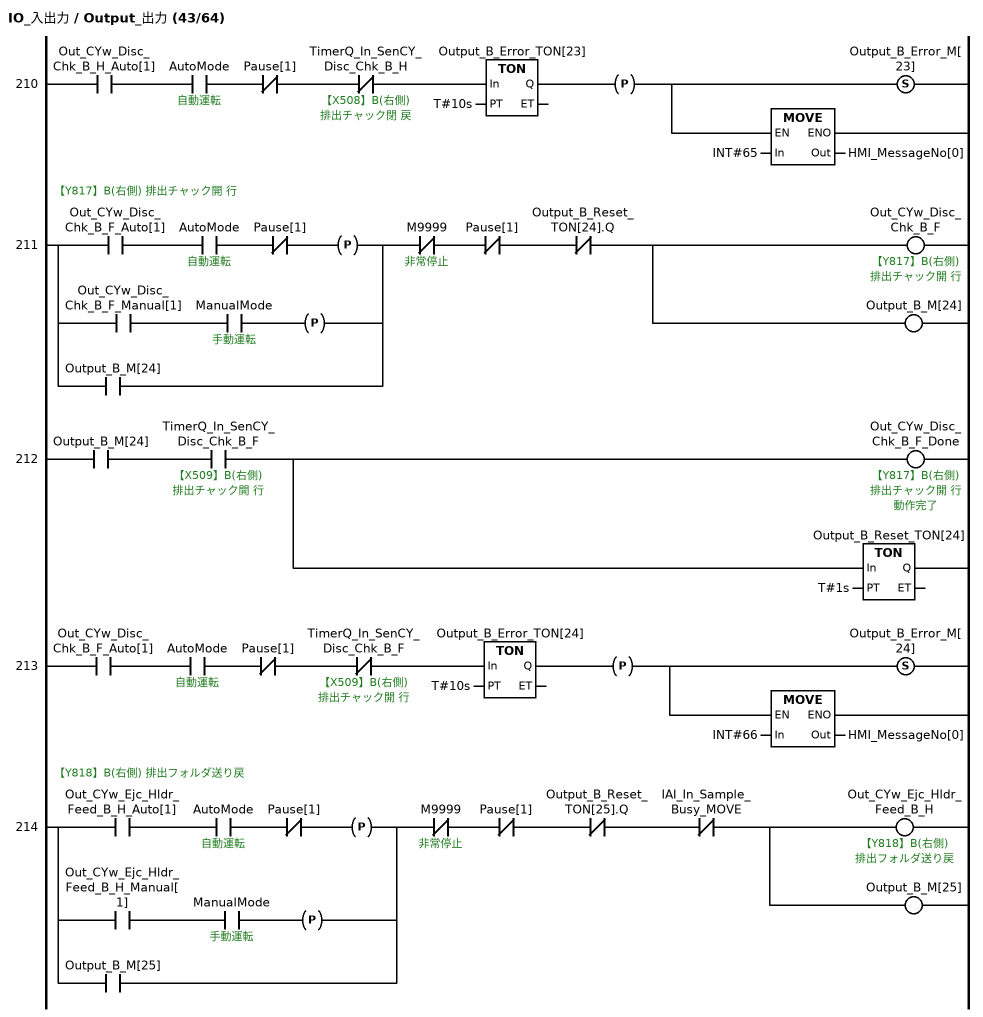
(* Rung 210 *)
Output_B_Error_TON[23](In := Out_CYw_Disc_Chk_B_H_Auto[1] AND AutoMode AND NOT Pause[1] AND NOT TimerQ_In_SenCY_Disc_Chk_B_H, PT := T#10s);
_e308(CLK := Output_B_Error_TON[23].Q);
IF _e308.Q THEN
    Output_B_Error_M[23] := TRUE;
    HMI_MessageNo[0] := INT#65;
END_IF;
(* Rung 211: 【Y817】B(右側) 排出チャック開 行 *)
_e309(CLK := Out_CYw_Disc_Chk_B_F_Auto[1] AND AutoMode AND NOT Pause[1]);
_e310(CLK := Out_CYw_Disc_Chk_B_F_Manual[1] AND ManualMode);
_p311 := (_e309.Q OR _e310.Q OR Output_B_M[24]) AND NOT M9999 AND NOT Pause[1] AND NOT Output_B_Reset_TON[24].Q;
Out_CYw_Disc_Chk_B_F := _p311;
Output_B_M[24] := _p311;
(* Rung 212 *)
Out_CYw_Disc_Chk_B_F_Done := Output_B_M[24] AND TimerQ_In_SenCY_Disc_Chk_B_F;
Output_B_Reset_TON[24](In := Output_B_M[24] AND TimerQ_In_SenCY_Disc_Chk_B_F, PT := T#1s);
(* Rung 213 *)
Output_B_Error_TON[24](In := Out_CYw_Disc_Chk_B_F_Auto[1] AND AutoMode AND NOT Pause[1] AND NOT TimerQ_In_SenCY_Disc_Chk_B_F, PT := T#10s);
_e312(CLK := Output_B_Error_TON[24].Q);
IF _e312.Q THEN
    Output_B_Error_M[24] := TRUE;
    HMI_MessageNo[0] := INT#66;
END_IF;
(* Rung 214: 【Y818】B(右側) 排出フォルダ送り戻 *)
_e313(CLK := Out_CYw_Ejc_Hldr_Feed_B_H_Auto[1] AND AutoMode AND NOT Pause[1]);
_e314(CLK := Out_CYw_Ejc_Hldr_Feed_B_H_Manual[1] AND ManualMode);
_p315 := (_e313.Q OR _e314.Q OR Output_B_M[25]) AND NOT M9999 AND NOT Pause[1] AND NOT Output_B_Reset_TON[25].Q AND NOT IAI_In_Sample_Busy_MOVE;
Out_CYw_Ejc_Hldr_Feed_B_H := _p315;
Output_B_M[25] := _p315;

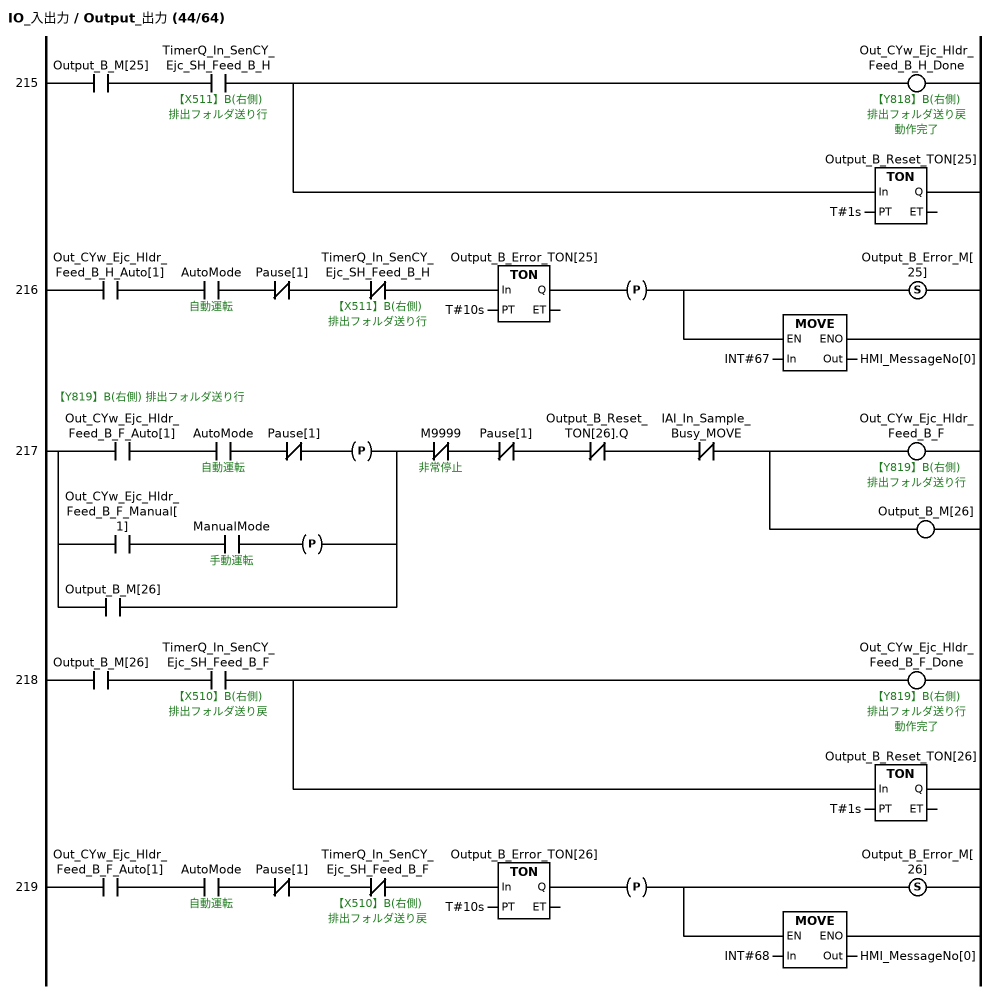
(* Rung 215 *)
_p316 := Output_B_M[25] AND TimerQ_In_SenCY_Ejc_SH_Feed_B_H;
Out_CYw_Ejc_Hldr_Feed_B_H_Done := _p316;
Output_B_Reset_TON[25](In := _p316, PT := T#1s);
(* Rung 216 *)
Output_B_Error_TON[25](In := Out_CYw_Ejc_Hldr_Feed_B_H_Auto[1] AND AutoMode AND NOT Pause[1] AND NOT TimerQ_In_SenCY_Ejc_SH_Feed_B_H, PT := T#10s);
_e317(CLK := Output_B_Error_TON[25].Q);
IF _e317.Q THEN
    Output_B_Error_M[25] := TRUE;
    HMI_MessageNo[0] := INT#67;
END_IF;
(* Rung 217: 【Y819】B(右側) 排出フォルダ送り行 *)
_e318(CLK := Out_CYw_Ejc_Hldr_Feed_B_F_Auto[1] AND AutoMode AND NOT Pause[1]);
_e319(CLK := Out_CYw_Ejc_Hldr_Feed_B_F_Manual[1] AND ManualMode);
_p320 := (_e318.Q OR _e319.Q OR Output_B_M[26]) AND NOT M9999 AND NOT Pause[1] AND NOT Output_B_Reset_TON[26].Q AND NOT IAI_In_Sample_Busy_MOVE;
Out_CYw_Ejc_Hldr_Feed_B_F := _p320;
Output_B_M[26] := _p320;
(* Rung 218 *)
_p321 := Output_B_M[26] AND TimerQ_In_SenCY_Ejc_SH_Feed_B_F;
Out_CYw_Ejc_Hldr_Feed_B_F_Done := _p321;
Output_B_Reset_TON[26](In := _p321, PT := T#1s);
(* Rung 219 *)
Output_B_Error_TON[26](In := Out_CYw_Ejc_Hldr_Feed_B_F_Auto[1] AND AutoMode AND NOT Pause[1] AND NOT TimerQ_In_SenCY_Ejc_SH_Feed_B_F, PT := T#10s);
_e322(CLK := Output_B_Error_TON[26].Q);
IF _e322.Q THEN
    Output_B_Error_M[26] := TRUE;
    HMI_MessageNo[0] := INT#68;
END_IF;

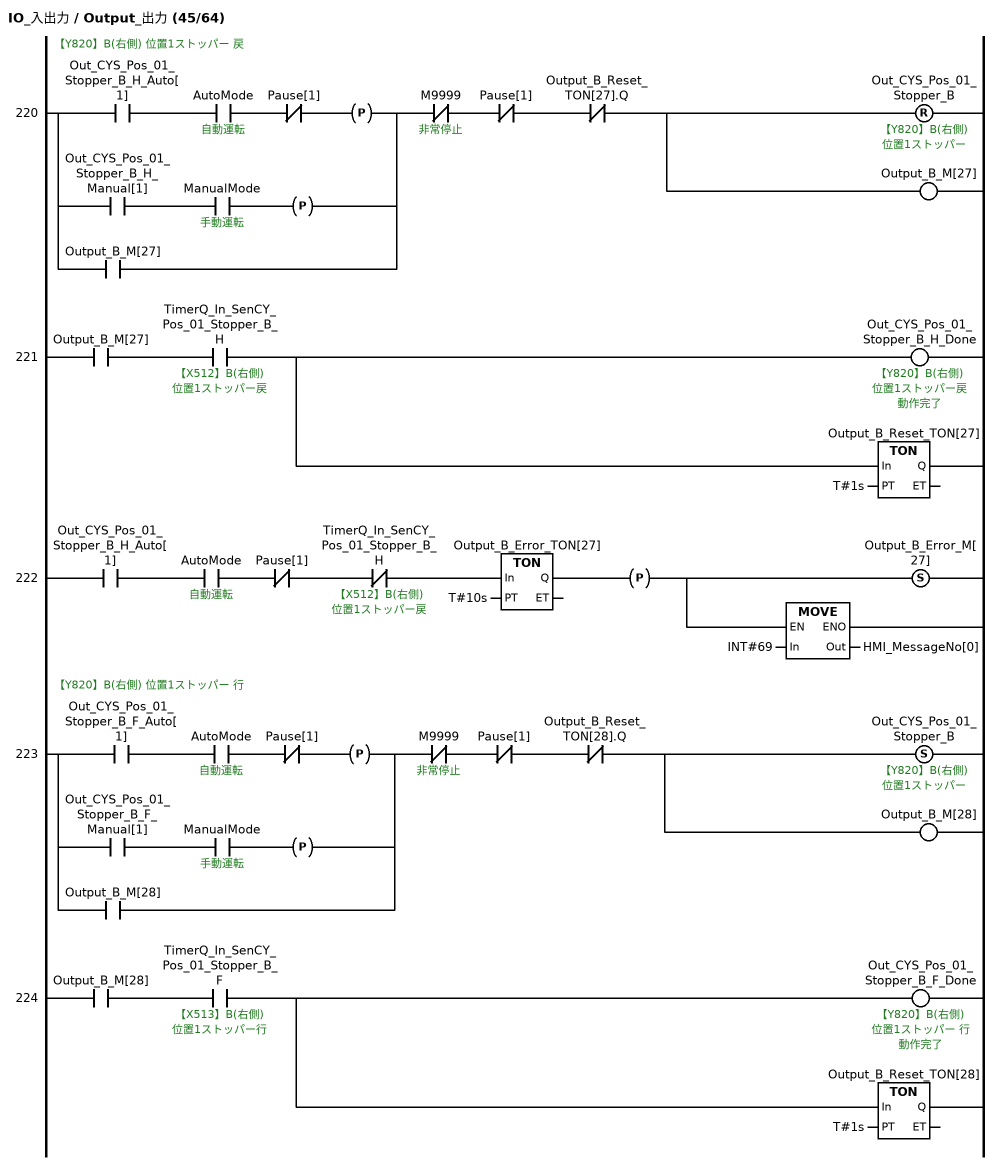
(* Rung 220: 【Y820】B(右側) 位置1ストッパー 戻 *)
_e323(CLK := Out_CYS_Pos_01_Stopper_B_H_Auto[1] AND AutoMode AND NOT Pause[1]);
_e324(CLK := Out_CYS_Pos_01_Stopper_B_H_Manual[1] AND ManualMode);
_p325 := (_e323.Q OR _e324.Q OR Output_B_M[27]) AND NOT M9999 AND NOT Pause[1] AND NOT Output_B_Reset_TON[27].Q;
IF _p325 THEN Out_CYS_Pos_01_Stopper_B := FALSE; END_IF;
Output_B_M[27] := _p325;
(* Rung 221 *)
_p326 := Output_B_M[27] AND TimerQ_In_SenCY_Pos_01_Stopper_B_H;
Out_CYS_Pos_01_Stopper_B_H_Done := _p326;
Output_B_Reset_TON[27](In := _p326, PT := T#1s);
(* Rung 222 *)
Output_B_Error_TON[27](In := Out_CYS_Pos_01_Stopper_B_H_Auto[1] AND AutoMode AND NOT Pause[1] AND NOT TimerQ_In_SenCY_Pos_01_Stopper_B_H, PT := T#10s);
_e327(CLK := Output_B_Error_TON[27].Q);
IF _e327.Q THEN
    Output_B_Error_M[27] := TRUE;
    HMI_MessageNo[0] := INT#69;
END_IF;
(* Rung 223: 【Y820】B(右側) 位置1ストッパー 行 *)
_e328(CLK := Out_CYS_Pos_01_Stopper_B_F_Auto[1] AND AutoMode AND NOT Pause[1]);
_e329(CLK := Out_CYS_Pos_01_Stopper_B_F_Manual[1] AND ManualMode);
_p330 := (_e328.Q OR _e329.Q OR Output_B_M[28]) AND NOT M9999 AND NOT Pause[1] AND NOT Output_B_Reset_TON[28].Q;
IF _p330 THEN Out_CYS_Pos_01_Stopper_B := TRUE; END_IF;
Output_B_M[28] := _p330;
(* Rung 224 *)
_p331 := Output_B_M[28] AND TimerQ_In_SenCY_Pos_01_Stopper_B_F;
Out_CYS_Pos_01_Stopper_B_F_Done := _p331;
Output_B_Reset_TON[28](In := _p331, PT := T#1s);

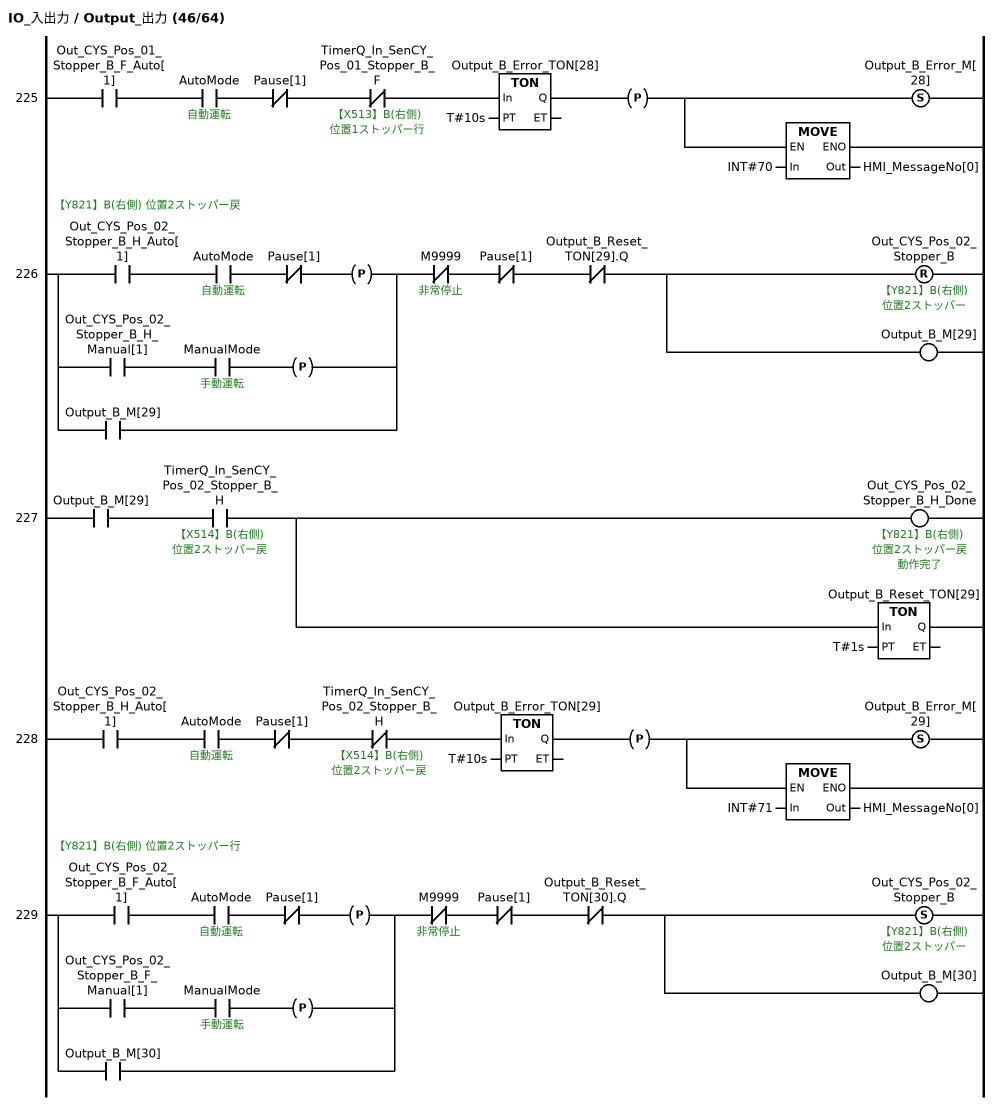
(* Rung 225 *)
Output_B_Error_TON[28](In := Out_CYS_Pos_01_Stopper_B_F_Auto[1] AND AutoMode AND NOT Pause[1] AND NOT TimerQ_In_SenCY_Pos_01_Stopper_B_F, PT := T#10s);
_e332(CLK := Output_B_Error_TON[28].Q);
IF _e332.Q THEN
    Output_B_Error_M[28] := TRUE;
    HMI_MessageNo[0] := INT#70;
END_IF;
(* Rung 226: 【Y821】B(右側) 位置2ストッパー戻 *)
_e333(CLK := Out_CYS_Pos_02_Stopper_B_H_Auto[1] AND AutoMode AND NOT Pause[1]);
_e334(CLK := Out_CYS_Pos_02_Stopper_B_H_Manual[1] AND ManualMode);
_p335 := (_e333.Q OR _e334.Q OR Output_B_M[29]) AND NOT M9999 AND NOT Pause[1] AND NOT Output_B_Reset_TON[29].Q;
IF _p335 THEN Out_CYS_Pos_02_Stopper_B := FALSE; END_IF;
Output_B_M[29] := _p335;
(* Rung 227 *)
_p336 := Output_B_M[29] AND TimerQ_In_SenCY_Pos_02_Stopper_B_H;
Out_CYS_Pos_02_Stopper_B_H_Done := _p336;
Output_B_Reset_TON[29](In := _p336, PT := T#1s);
(* Rung 228 *)
Output_B_Error_TON[29](In := Out_CYS_Pos_02_Stopper_B_H_Auto[1] AND AutoMode AND NOT Pause[1] AND NOT TimerQ_In_SenCY_Pos_02_Stopper_B_H, PT := T#10s);
_e337(CLK := Output_B_Error_TON[29].Q);
IF _e337.Q THEN
    Output_B_Error_M[29] := TRUE;
    HMI_MessageNo[0] := INT#71;
END_IF;
(* Rung 229: 【Y821】B(右側) 位置2ストッパー行 *)
_e338(CLK := Out_CYS_Pos_02_Stopper_B_F_Auto[1] AND AutoMode AND NOT Pause[1]);
_e339(CLK := Out_CYS_Pos_02_Stopper_B_F_Manual[1] AND ManualMode);
_p340 := (_e338.Q OR _e339.Q OR Output_B_M[30]) AND NOT M9999 AND NOT Pause[1] AND NOT Output_B_Reset_TON[30].Q;
IF _p340 THEN Out_CYS_Pos_02_Stopper_B := TRUE; END_IF;
Output_B_M[30] := _p340;

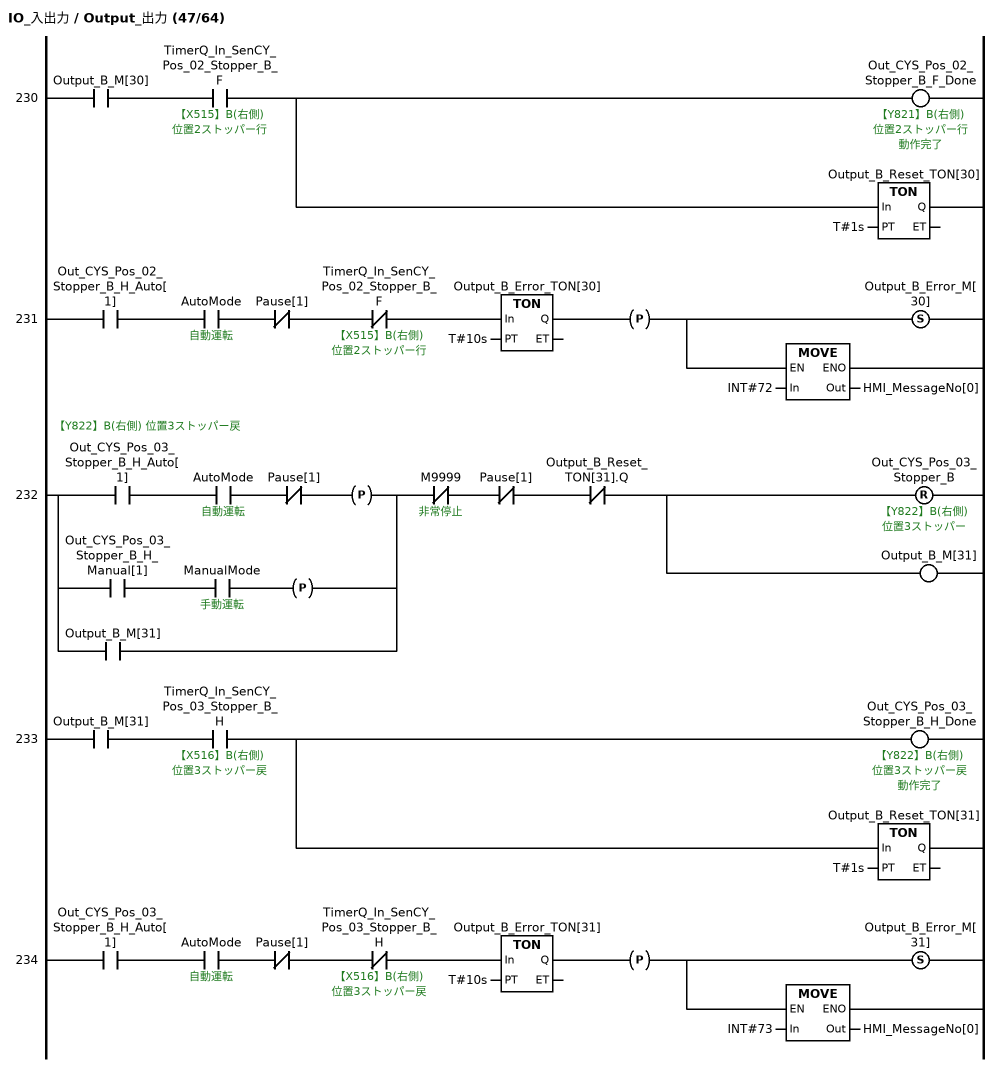
(* Rung 230 *)
_p341 := Output_B_M[30] AND TimerQ_In_SenCY_Pos_02_Stopper_B_F;
Out_CYS_Pos_02_Stopper_B_F_Done := _p341;
Output_B_Reset_TON[30](In := _p341, PT := T#1s);
(* Rung 231 *)
Output_B_Error_TON[30](In := Out_CYS_Pos_02_Stopper_B_H_Auto[1] AND AutoMode AND NOT Pause[1] AND NOT TimerQ_In_SenCY_Pos_02_Stopper_B_F, PT := T#10s);
_e342(CLK := Output_B_Error_TON[30].Q);
IF _e342.Q THEN
    Output_B_Error_M[30] := TRUE;
    HMI_MessageNo[0] := INT#72;
END_IF;
(* Rung 232: 【Y822】B(右側) 位置3ストッパー戻 *)
_e343(CLK := Out_CYS_Pos_03_Stopper_B_H_Auto[1] AND AutoMode AND NOT Pause[1]);
_e344(CLK := Out_CYS_Pos_03_Stopper_B_H_Manual[1] AND ManualMode);
_p345 := (_e343.Q OR _e344.Q OR Output_B_M[31]) AND NOT M9999 AND NOT Pause[1] AND NOT Output_B_Reset_TON[31].Q;
IF _p345 THEN Out_CYS_Pos_03_Stopper_B := FALSE; END_IF;
Output_B_M[31] := _p345;
(* Rung 233 *)
_p346 := Output_B_M[31] AND TimerQ_In_SenCY_Pos_03_Stopper_B_H;
Out_CYS_Pos_03_Stopper_B_H_Done := _p346;
Output_B_Reset_TON[31](In := _p346, PT := T#1s);
(* Rung 234 *)
Output_B_Error_TON[31](In := Out_CYS_Pos_03_Stopper_B_H_Auto[1] AND AutoMode AND NOT Pause[1] AND NOT TimerQ_In_SenCY_Pos_03_Stopper_B_H, PT := T#10s);
_e347(CLK := Output_B_Error_TON[31].Q);
IF _e347.Q THEN
    Output_B_Error_M[31] := TRUE;
    HMI_MessageNo[0] := INT#73;
END_IF;

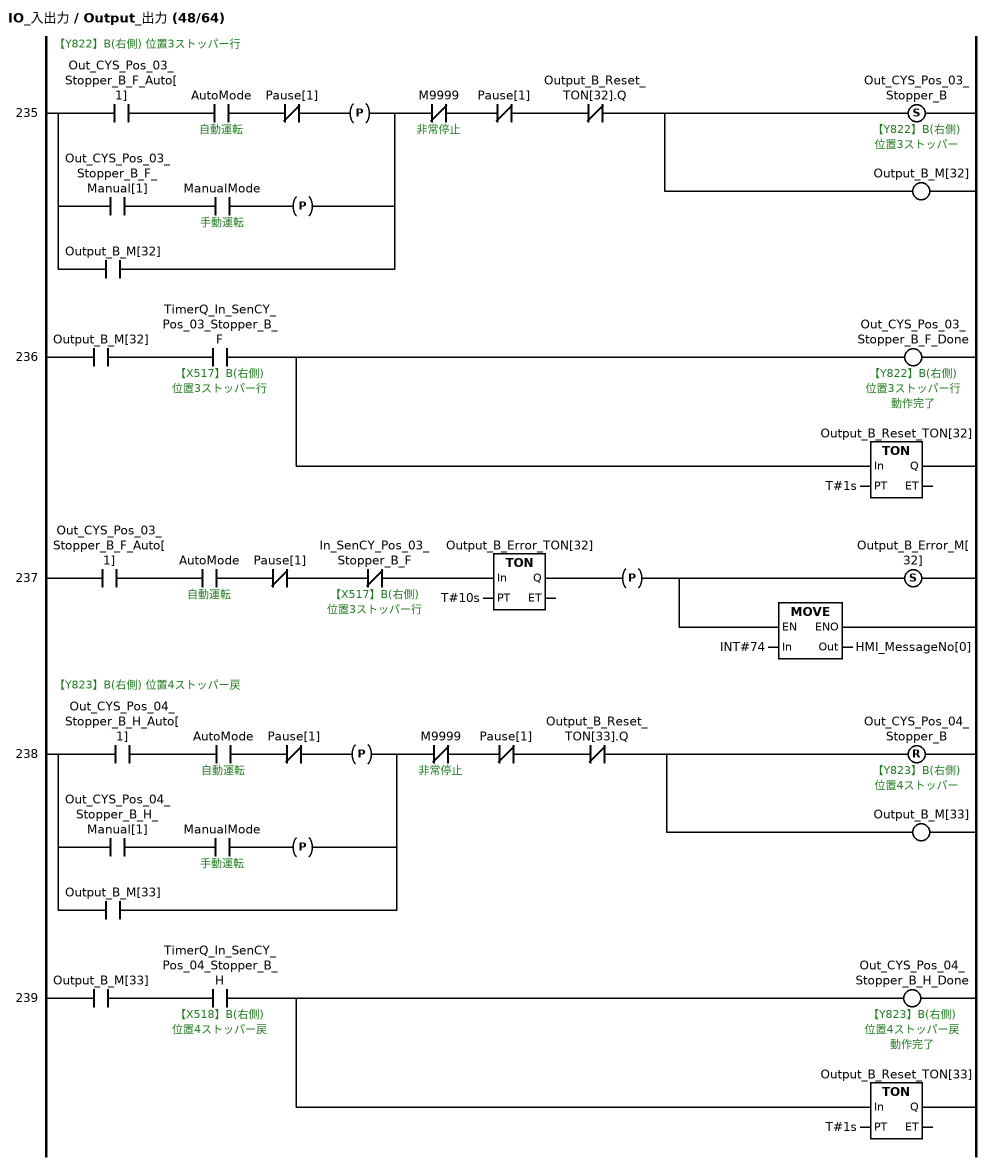
(* Rung 235: 【Y822】B(右側) 位置3ストッパー行 *)
_e348(CLK := Out_CYS_Pos_03_Stopper_B_F_Auto[1] AND AutoMode AND NOT Pause[1]);
_e349(CLK := Out_CYS_Pos_03_Stopper_B_F_Manual[1] AND ManualMode);
_p350 := (_e348.Q OR _e349.Q OR Output_B_M[32]) AND NOT M9999 AND NOT Pause[1] AND NOT Output_B_Reset_TON[32].Q;
IF _p350 THEN Out_CYS_Pos_03_Stopper_B := TRUE; END_IF;
Output_B_M[32] := _p350;
(* Rung 236 *)
_p351 := Output_B_M[32] AND TimerQ_In_SenCY_Pos_03_Stopper_B_F;
Out_CYS_Pos_03_Stopper_B_F_Done := _p351;
Output_B_Reset_TON[32](In := _p351, PT := T#1s);
(* Rung 237 *)
Output_B_Error_TON[32](In := Out_CYS_Pos_03_Stopper_B_F_Auto[1] AND AutoMode AND NOT Pause[1] AND NOT In_SenCY_Pos_03_Stopper_B_F, PT := T#10s);
_e352(CLK := Output_B_Error_TON[32].Q);
IF _e352.Q THEN
    Output_B_Error_M[32] := TRUE;
    HMI_MessageNo[0] := INT#74;
END_IF;
(* Rung 238: 【Y823】B(右側) 位置4ストッパー戻 *)
_e353(CLK := Out_CYS_Pos_04_Stopper_B_H_Auto[1] AND AutoMode AND NOT Pause[1]);
_e354(CLK := Out_CYS_Pos_04_Stopper_B_H_Manual[1] AND ManualMode);
_p355 := (_e353.Q OR _e354.Q OR Output_B_M[33]) AND NOT M9999 AND NOT Pause[1] AND NOT Output_B_Reset_TON[33].Q;
IF _p355 THEN Out_CYS_Pos_04_Stopper_B := FALSE; END_IF;
Output_B_M[33] := _p355;
(* Rung 239 *)
_p356 := Output_B_M[33] AND TimerQ_In_SenCY_Pos_04_Stopper_B_H;
Out_CYS_Pos_04_Stopper_B_H_Done := _p356;
Output_B_Reset_TON[33](In := _p356, PT := T#1s);

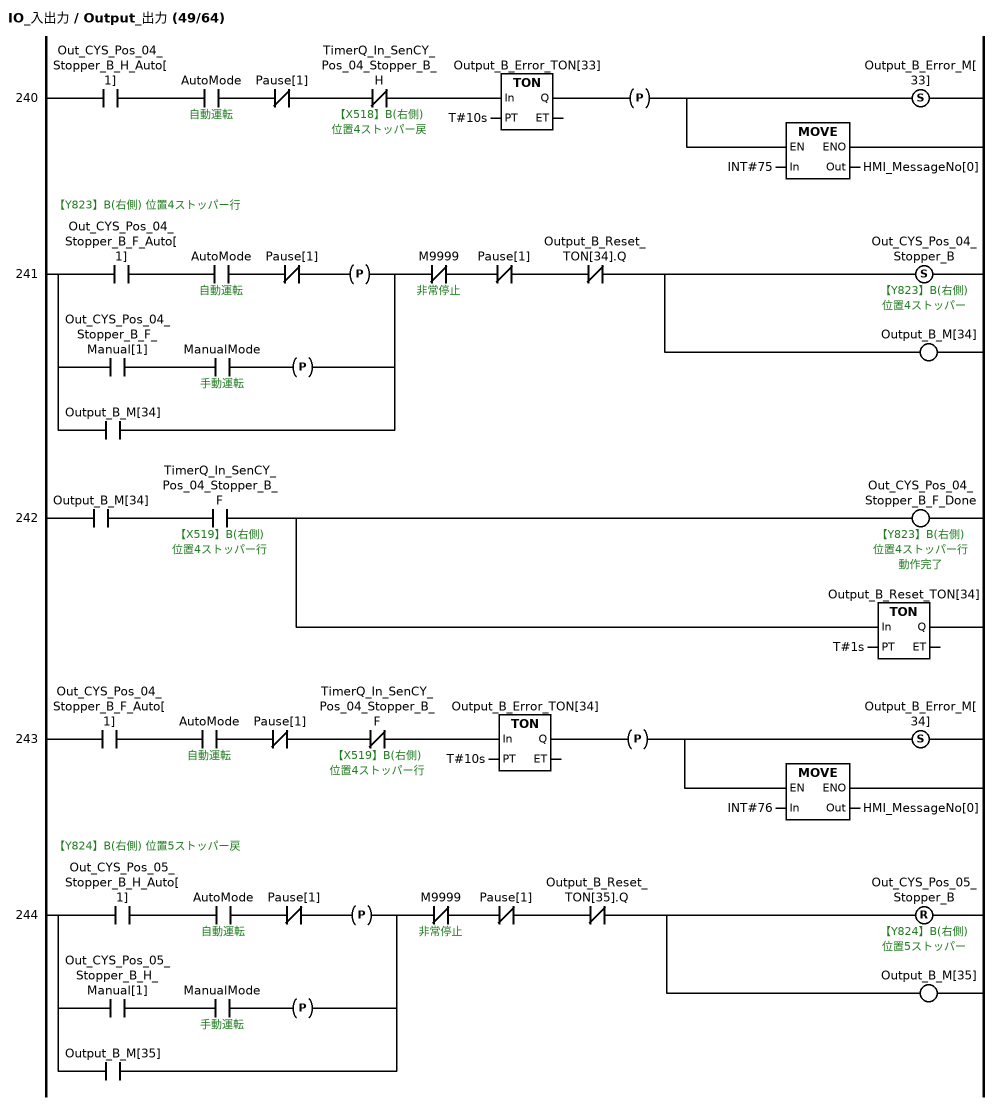
(* Rung 240 *)
Output_B_Error_TON[33](In := Out_CYS_Pos_04_Stopper_B_H_Auto[1] AND AutoMode AND NOT Pause[1] AND NOT TimerQ_In_SenCY_Pos_04_Stopper_B_H, PT := T#10s);
_e357(CLK := Output_B_Error_TON[33].Q);
IF _e357.Q THEN
    Output_B_Error_M[33] := TRUE;
    HMI_MessageNo[0] := INT#75;
END_IF;
(* Rung 241: 【Y823】B(右側) 位置4ストッパー行 *)
_e358(CLK := Out_CYS_Pos_04_Stopper_B_F_Auto[1] AND AutoMode AND NOT Pause[1]);
_e359(CLK := Out_CYS_Pos_04_Stopper_B_F_Manual[1] AND ManualMode);
_p360 := (_e358.Q OR _e359.Q OR Output_B_M[34]) AND NOT M9999 AND NOT Pause[1] AND NOT Output_B_Reset_TON[34].Q;
IF _p360 THEN Out_CYS_Pos_04_Stopper_B := TRUE; END_IF;
Output_B_M[34] := _p360;
(* Rung 242 *)
_p361 := Output_B_M[34] AND TimerQ_In_SenCY_Pos_04_Stopper_B_F;
Out_CYS_Pos_04_Stopper_B_F_Done := _p361;
Output_B_Reset_TON[34](In := _p361, PT := T#1s);
(* Rung 243 *)
Output_B_Error_TON[34](In := Out_CYS_Pos_04_Stopper_B_F_Auto[1] AND AutoMode AND NOT Pause[1] AND NOT TimerQ_In_SenCY_Pos_04_Stopper_B_F, PT := T#10s);
_e362(CLK := Output_B_Error_TON[34].Q);
IF _e362.Q THEN
    Output_B_Error_M[34] := TRUE;
    HMI_MessageNo[0] := INT#76;
END_IF;
(* Rung 244: 【Y824】B(右側) 位置5ストッパー戻 *)
_e363(CLK := Out_CYS_Pos_05_Stopper_B_H_Auto[1] AND AutoMode AND NOT Pause[1]);
_e364(CLK := Out_CYS_Pos_05_Stopper_B_H_Manual[1] AND ManualMode);
_p365 := (_e363.Q OR _e364.Q OR Output_B_M[35]) AND NOT M9999 AND NOT Pause[1] AND NOT Output_B_Reset_TON[35].Q;
IF _p365 THEN Out_CYS_Pos_05_Stopper_B := FALSE; END_IF;
Output_B_M[35] := _p365;

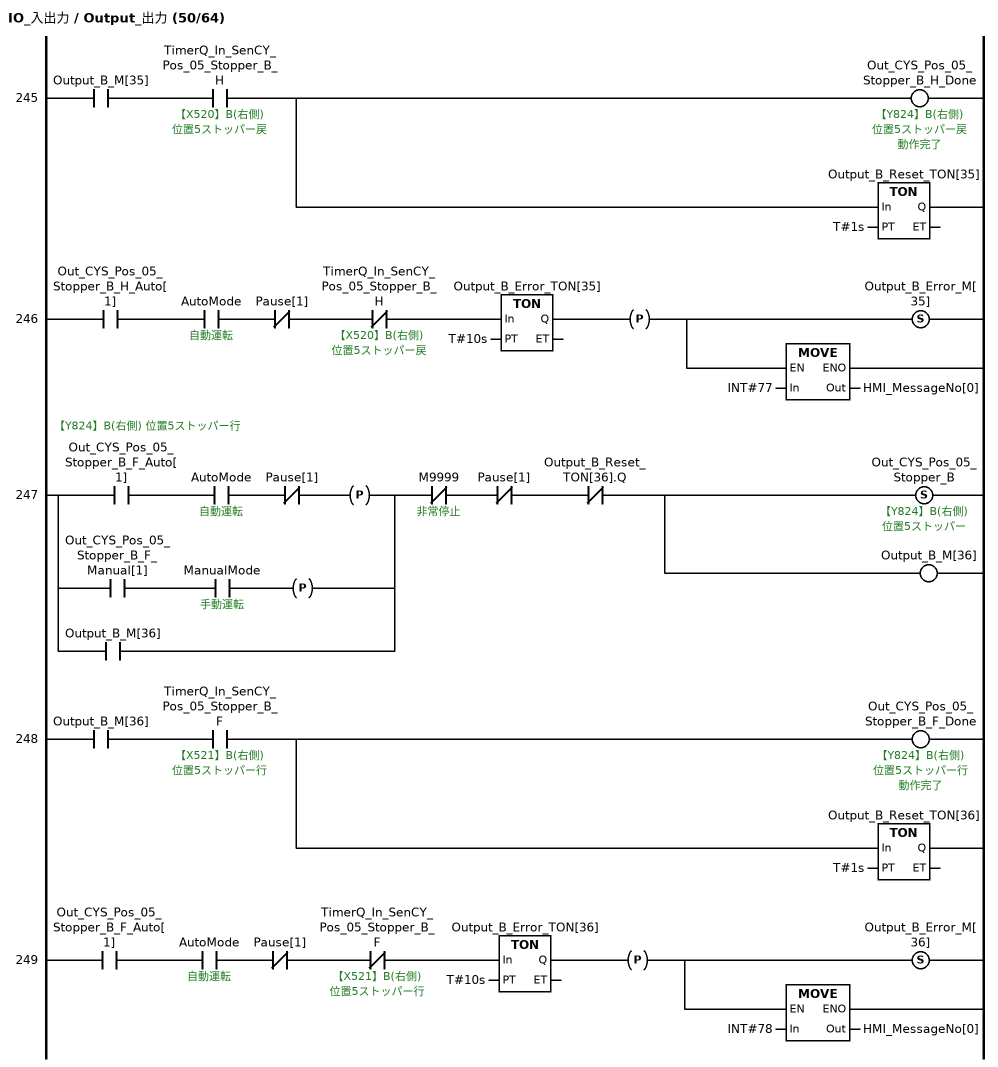
(* Rung 245 *)
_p366 := Output_B_M[35] AND TimerQ_In_SenCY_Pos_05_Stopper_B_H;
Out_CYS_Pos_05_Stopper_B_H_Done := _p366;
Output_B_Reset_TON[35](In := _p366, PT := T#1s);
(* Rung 246 *)
Output_B_Error_TON[35](In := Out_CYS_Pos_05_Stopper_B_H_Auto[1] AND AutoMode AND NOT Pause[1] AND NOT TimerQ_In_SenCY_Pos_05_Stopper_B_H, PT := T#10s);
_e367(CLK := Output_B_Error_TON[35].Q);
IF _e367.Q THEN
    Output_B_Error_M[35] := TRUE;
    HMI_MessageNo[0] := INT#77;
END_IF;
(* Rung 247: 【Y824】B(右側) 位置5ストッパー行 *)
_e368(CLK := Out_CYS_Pos_05_Stopper_B_F_Auto[1] AND AutoMode AND NOT Pause[1]);
_e369(CLK := Out_CYS_Pos_05_Stopper_B_F_Manual[1] AND ManualMode);
_p370 := (_e368.Q OR _e369.Q OR Output_B_M[36]) AND NOT M9999 AND NOT Pause[1] AND NOT Output_B_Reset_TON[36].Q;
IF _p370 THEN Out_CYS_Pos_05_Stopper_B := TRUE; END_IF;
Output_B_M[36] := _p370;
(* Rung 248 *)
_p371 := Output_B_M[36] AND TimerQ_In_SenCY_Pos_05_Stopper_B_F;
Out_CYS_Pos_05_Stopper_B_F_Done := _p371;
Output_B_Reset_TON[36](In := _p371, PT := T#1s);
(* Rung 249 *)
Output_B_Error_TON[36](In := Out_CYS_Pos_05_Stopper_B_F_Auto[1] AND AutoMode AND NOT Pause[1] AND NOT TimerQ_In_SenCY_Pos_05_Stopper_B_F, PT := T#10s);
_e372(CLK := Output_B_Error_TON[36].Q);
IF _e372.Q THEN
    Output_B_Error_M[36] := TRUE;
    HMI_MessageNo[0] := INT#78;
END_IF;

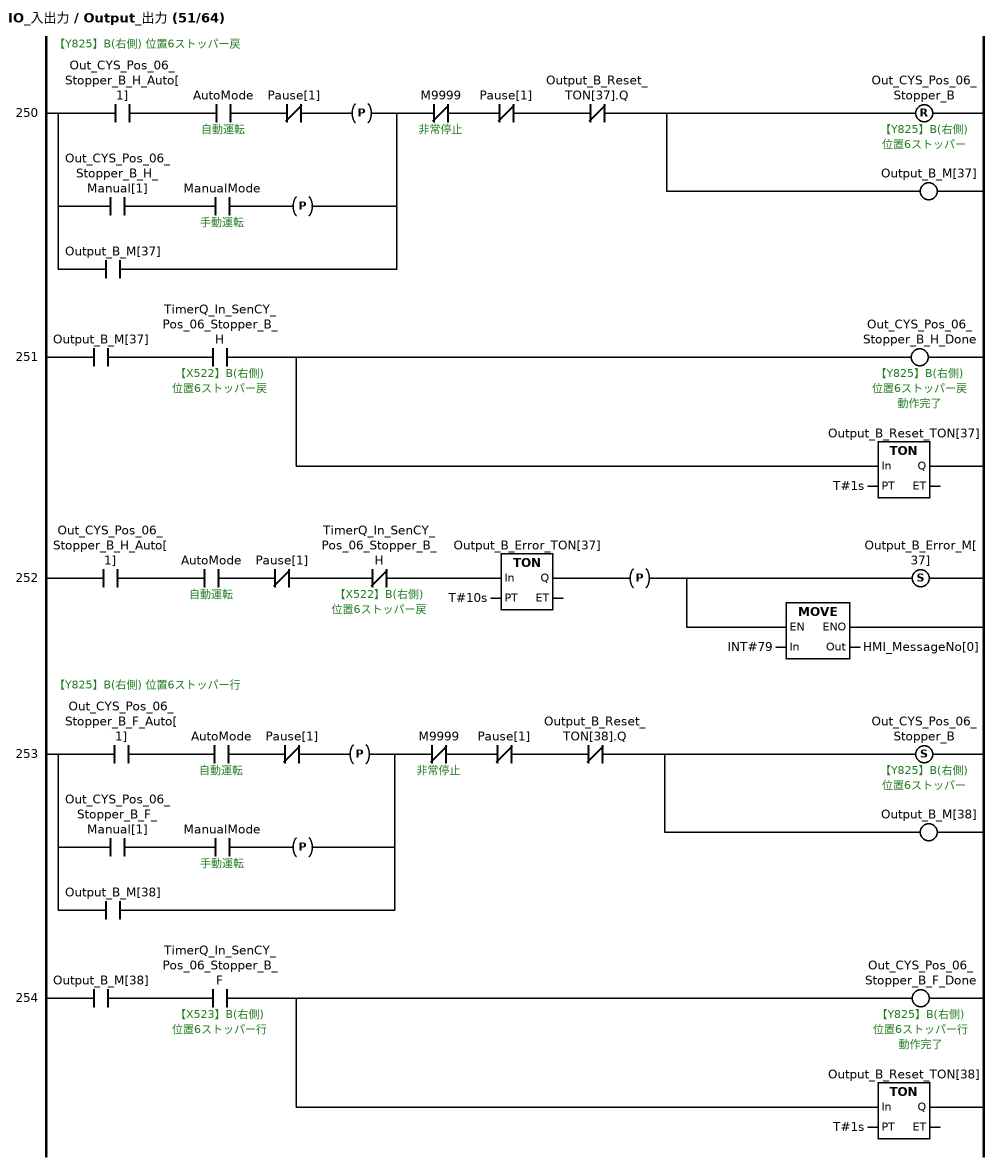
(* Rung 250: 【Y825】B(右側) 位置6ストッパー戻 *)
_e373(CLK := Out_CYS_Pos_06_Stopper_B_H_Auto[1] AND AutoMode AND NOT Pause[1]);
_e374(CLK := Out_CYS_Pos_06_Stopper_B_H_Manual[1] AND ManualMode);
_p375 := (_e373.Q OR _e374.Q OR Output_B_M[37]) AND NOT M9999 AND NOT Pause[1] AND NOT Output_B_Reset_TON[37].Q;
IF _p375 THEN Out_CYS_Pos_06_Stopper_B := FALSE; END_IF;
Output_B_M[37] := _p375;
(* Rung 251 *)
_p376 := Output_B_M[37] AND TimerQ_In_SenCY_Pos_06_Stopper_B_H;
Out_CYS_Pos_06_Stopper_B_H_Done := _p376;
Output_B_Reset_TON[37](In := _p376, PT := T#1s);
(* Rung 252 *)
Output_B_Error_TON[37](In := Out_CYS_Pos_06_Stopper_B_H_Auto[1] AND AutoMode AND NOT Pause[1] AND NOT TimerQ_In_SenCY_Pos_06_Stopper_B_H, PT := T#10s);
_e377(CLK := Output_B_Error_TON[37].Q);
IF _e377.Q THEN
    Output_B_Error_M[37] := TRUE;
    HMI_MessageNo[0] := INT#79;
END_IF;
(* Rung 253: 【Y825】B(右側) 位置6ストッパー行 *)
_e378(CLK := Out_CYS_Pos_06_Stopper_B_F_Auto[1] AND AutoMode AND NOT Pause[1]);
_e379(CLK := Out_CYS_Pos_06_Stopper_B_F_Manual[1] AND ManualMode);
_p380 := (_e378.Q OR _e379.Q OR Output_B_M[38]) AND NOT M9999 AND NOT Pause[1] AND NOT Output_B_Reset_TON[38].Q;
IF _p380 THEN Out_CYS_Pos_06_Stopper_B := TRUE; END_IF;
Output_B_M[38] := _p380;
(* Rung 254 *)
_p381 := Output_B_M[38] AND TimerQ_In_SenCY_Pos_06_Stopper_B_F;
Out_CYS_Pos_06_Stopper_B_F_Done := _p381;
Output_B_Reset_TON[38](In := _p381, PT := T#1s);

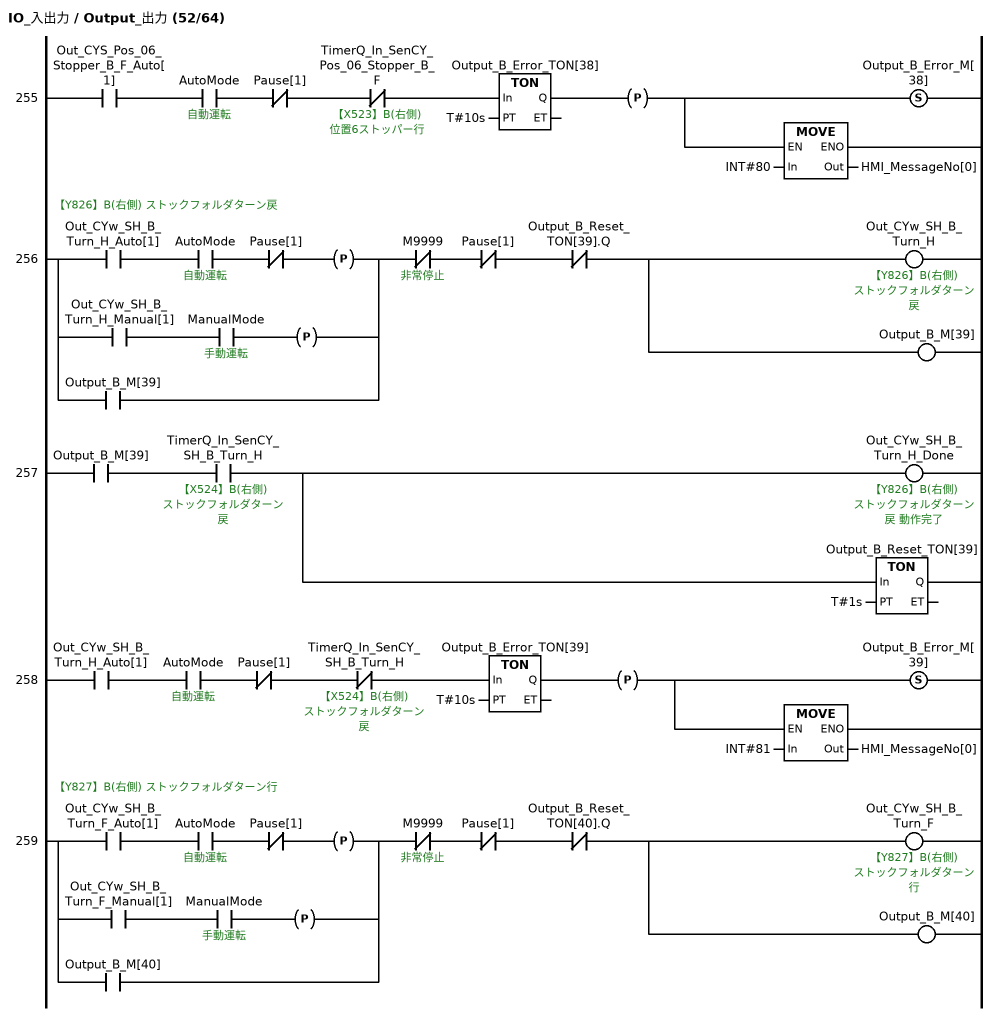
(* Rung 255 *)
Output_B_Error_TON[38](In := Out_CYS_Pos_06_Stopper_B_F_Auto[1] AND AutoMode AND NOT Pause[1] AND NOT TimerQ_In_SenCY_Pos_06_Stopper_B_F, PT := T#10s);
_e382(CLK := Output_B_Error_TON[38].Q);
IF _e382.Q THEN
    Output_B_Error_M[38] := TRUE;
    HMI_MessageNo[0] := INT#80;
END_IF;
(* Rung 256: 【Y826】B(右側) ストックフォルダターン戻 *)
_e383(CLK := Out_CYw_SH_B_Turn_H_Auto[1] AND AutoMode AND NOT Pause[1]);
_e384(CLK := Out_CYw_SH_B_Turn_H_Manual[1] AND ManualMode);
_p385 := (_e383.Q OR _e384.Q OR Output_B_M[39]) AND NOT M9999 AND NOT Pause[1] AND NOT Output_B_Reset_TON[39].Q;
Out_CYw_SH_B_Turn_H := _p385;
Output_B_M[39] := _p385;
(* Rung 257 *)
Out_CYw_SH_B_Turn_H_Done := Output_B_M[39] AND TimerQ_In_SenCY_SH_B_Turn_H;
Output_B_Reset_TON[39](In := Output_B_M[39] AND TimerQ_In_SenCY_SH_B_Turn_H, PT := T#1s);
(* Rung 258 *)
Output_B_Error_TON[39](In := Out_CYw_SH_B_Turn_H_Auto[1] AND AutoMode AND NOT Pause[1] AND NOT TimerQ_In_SenCY_SH_B_Turn_H, PT := T#10s);
_e386(CLK := Output_B_Error_TON[39].Q);
IF _e386.Q THEN
    Output_B_Error_M[39] := TRUE;
    HMI_MessageNo[0] := INT#81;
END_IF;
(* Rung 259: 【Y827】B(右側) ストックフォルダターン行 *)
_e387(CLK := Out_CYw_SH_B_Turn_F_Auto[1] AND AutoMode AND NOT Pause[1]);
_e388(CLK := Out_CYw_SH_B_Turn_F_Manual[1] AND ManualMode);
_p389 := (_e387.Q OR _e388.Q OR Output_B_M[40]) AND NOT M9999 AND NOT Pause[1] AND NOT Output_B_Reset_TON[40].Q;
Out_CYw_SH_B_Turn_F := _p389;
Output_B_M[40] := _p389;

